(* IEC 61131-3 sources: daoli-st-library/DL_MathData (part 28) *)

(* ---- FC_DL_WordToBytes.st ---- *)
(*==============================================================================
 * 组件名称 (Component)  : FC_DL_WordToBytes
 * 所属子库 (Sublibrary) : DL_MathData
 * 当前版本 (Version)    : 1.0.0
 * 兼容性   (Platform)   : CODESYS 3.5 / TwinCAT 3 / 汇川 InoProShop / Machine Expert
 *                         仅依赖 Standard.library（SHR / AND / 类型转换），零厂商方言
 * 来源标签 (Source)     : t2-1-lgf-converter（字节序拆解族，clean-room 编写）
 * 功能描述 (Function)   : WORD / DWORD 按字节序拆解为 BYTE 数组（写经指针输出）。
 *                         槽位语义与 FC_DL_WordFromBytes 完全对偶：槽 0 = 最高字节；
 *                         映射为对合映射（ involutive），同一序号下
 *                         WordToBytes(WordFromBytes(bytes, eOrder, len), eOrder, len)
 *                         逐字节还原源数组（round-trip 验收）。
 *                         nValueLen = 2 时只取低 16 位（高 16 位忽略）。
 *                         缓冲长度不足时钳位只写前 nBufLen 个槽位并置信息级。
 * 归属声明 (Ownership)  : E_DL_ByteOrder 归属 DL_MathData\FC_DL_SwapBytes32.st，
 *                         本件只引用不重声明（FB51-7）。
 * 边界与语义披露 (Boundary disclosure) :
 *   1) 指针 NIL 或缓冲长度 <= 0：结构性早退，不写任何字节，返回 FALSE（零写入语义）。
 *   2) 缓冲长度大于目标长度：多余槽位不触碰（不置码——缓冲边界由调用方持有，
 *      可观测性在调用方，R90 反证成立不加码）。
 *   3) 还原方向不饱和（R81 披露）：本件是拆解不是还原时刻 / 标识，拆解失败
 *      返回 FALSE + 故障级码，绝无静默饱和写入。
 *   4) 移位量上界 (nLenUse-1-j)*8 结构性 <= 24 < 32（DWORD 位宽），禁 MOD 归一的
 *      不变量由本披露承担（R48 口径）。
 *   5) 验收向量（与 FromBytes 对拍）：CDAB 序 16#0000_1234 -> {16#34, 16#12}；
 *      ABCD 16#1234_5678 -> {16#12,16#34,16#56,16#78}；缓冲 1 字节拆 DWORD
 *      -> 只写最高字节 + 信息级钳位。
 * 故障码表 (Error codes) :
 *   16#0001_03F5 [故障级] 缓冲指针 NIL 或 nBufLen <= 0，不写任何字节，返回 FALSE
 *                 反证：未写缓冲与「缓冲区内容本来如此」不可区分（本件无权回读
 *                 调用方缓冲），码位是唯一的失败事实出口。
 *   16#0001_03F6 [故障级] 字节序枚举越界（非 0..3），回退默认大端 eAbcd 继续服务
 *                 反证：回退结果与显式填 eAbcd 输出组合相同，码位承载组态有误事实。
 *   16#0001_04BA [信息级] 缓冲长度不足目标长度，已钳位只写前段
 *                 反证：钳位写入与「调用方只想要前段」输出组合相同，无码不可区分。
 *   16#0001_04BB [信息级] nValueLen 非 2/4，回退默认 WORD（2 字节）继续服务
 *                 反证：回退结果与显式填 2 相同，码位承载组态有误事实。
 * 码位总账 (Code ledger) : 16#0001_03F5 / 03F6 用 ｜ 16#0001_04BA / 04BB 用
 * 依赖     (Depends)    : TYPE E_DL_ByteOrder（属主 FC_DL_SwapBytes32.st，只引用）
 * 红线自检 (Redline)    : R1 ✓ 零全局变量与 VAR_EXTERNAL ｜ R2 ✓ 零 %I/%Q 物理地址
 *                         R3 ✓ 纯 IEC 61131-3（指针判空 + 标准移位/转换）
 *                         R4 ✓ 指针 NIL 闸 / 缓冲域闸 / 枚举域闸 / 全分支码位配对
 *                         R5 ✓ 全变量中英双语同行注释 ｜ R6 N/A（纯函数，无状态机）
 *                         R7 N/A（无定时器 / 边沿实例）
 * 修订历史 (Revision)   :
 *   2026-11-22  v1.0.0  首版入库（R68 构建轮 · 批 1 · 目标 5）
 *============================================================================*)
FUNCTION FC_DL_WordToBytes : BOOL
VAR_INPUT
    uValue    : DWORD;              // 待拆解值（WORD 目标时只取低 16 位）/ Value to split, low word only for WORD
    nValueLen : INT := 2;           // 值长度 [字节]，2 = WORD，4 = DWORD / Value length in bytes
    eOrder    : E_DL_ByteOrder;     // 字节序选择（属主 FC_DL_SwapBytes32.st）/ Byte order selector
    nBufLen   : INT;                // 输出缓冲长度 [字节]，<= 0 无效 / Output buffer length, <= 0 invalid
    pBuf      : POINTER TO BYTE;    // 输出缓冲首指针（指针本身不被改写，按输入口径）/ Output buffer pointer, never re-pointed
END_VAR
VAR_OUTPUT
    bWritten  : BOOL;    // 本拍写入成功 / Write succeeded this call
    bError    : BOOL;    // 故障标志（0307 / 0308 置位，R45 配对）/ Fault flag, set on 0307 and 0308
    uInfoId   : UDINT;   // 故障码，0 = 无故障（纯函数每拍重算）/ Error code, recomputed per call
END_VAR
VAR
    nWriteLen : INT;     // 本拍实际写入字节数 [个] / Bytes actually written this call
    nSlotByte : INT;     // 当前槽位映射回的源字节下标 / Byte index the current slot maps back to
    nShift    : DINT;    // 当前槽位移位量 [bit]，结构性 <= 24 / Slot shift amount
    uSlotVal  : DWORD;   // 当前槽位值（已掩码低 8 位）/ Current slot value, low 8 bits
    uB        : BYTE;    // 当前槽位字节 / Current slot byte
    nLenUse   : INT;     // 钳位后的值长度 [字节] / Clamped value length
    bOrderOk  : BOOL;    // 字节序枚举合法性 / Byte order validity
    j         : INT;     // 槽位遍历索引 / Slot loop index
END_VAR
VAR CONSTANT
    DL_WTB_LEN_MIN : INT      := 2;          // 值长度下限 [字节]（WORD）/ Value length floor, WORD
    DL_WTB_LEN_MAX : INT      := 4;          // 值长度上限 [字节]（DWORD）/ Value length ceiling, DWORD
    DL_WTB_MASK_FF : DWORD    := 16#0000_00FF; // 低 8 位掩码 / Low byte mask
END_VAR

(*------------------------------------------------------------------------------
 * 段 1｜安全预置（P-01 范式）：任何异常路径不写缓冲、返回 FALSE
 *      Safe preset: every exceptional path writes nothing and returns FALSE
 *-----------------------------------------------------------------------------*)
FC_DL_WordToBytes := FALSE;
bWritten := FALSE;
bError   := FALSE;
uInfoId  := 16#0000_0000;

(*------------------------------------------------------------------------------
 * 段 2｜域闸（R151 全枚举：指针 + 缓冲 + 值长度 + 枚举四闸）
 *      Domain gates: pointer, buffer, value length and enum
 *-----------------------------------------------------------------------------*)
IF (pBuf = 0) OR (nBufLen <= 0) THEN
    uInfoId := 16#0001_03F5;    // 故障级：指针 NIL 或缓冲非法 / Fault: NIL pointer or bad buffer
    bError  := TRUE;            // R45 配对 / Paired with the fault code
    RETURN;                     // 结构性早退：输出已全预置，零写入语义成立（规格明示豁免）
END_IF

IF (nValueLen < DL_WTB_LEN_MIN) OR (nValueLen > DL_WTB_LEN_MAX) THEN
    nLenUse := DL_WTB_LEN_MIN;  // 二级回退：钳回默认 WORD（R117 两级参数回退）
    uInfoId := 16#0001_04BB;    // 信息级：值长度非法回默认 / Info: length defaulted
ELSE
    nLenUse := nValueLen;       // 合法直通 / Valid pass-through
END_IF

bOrderOk := (eOrder = E_DL_ByteOrder.eAbcd) OR (eOrder = E_DL_ByteOrder.eDcba)
            OR (eOrder = E_DL_ByteOrder.eBadc) OR (eOrder = E_DL_ByteOrder.eCdab);
IF NOT bOrderOk THEN
    uInfoId := 16#0001_03F6;    // 故障级：字节序越界回默认大端（0142 风格先例口径）/ Fault: order defaulted
    bError  := TRUE;            // R45 配对 / Paired with the fault code
END_IF

(*------------------------------------------------------------------------------
 * 段 3｜写入长度钳位（边界 B4）：缓冲不足只写前段 + 信息级
 *      Write length clamp: short buffer writes the leading slots only
 *-----------------------------------------------------------------------------*)
IF nBufLen < nLenUse THEN
    nWriteLen := nBufLen;       // 钳位：只写缓冲能容纳的槽位 / Clamp to buffer capacity
    uInfoId   := 16#0001_04BA;  // 信息级：缓冲不足钳位 / Info: buffer clamped
ELSE
    nWriteLen := nLenUse;       // 充足：全量写入 / Full write
END_IF

(*------------------------------------------------------------------------------
 * 段 4｜拆解主体（边界 B1/B3）：取槽 -> 掩码 -> 降位 -> 反映射 -> 写缓冲
 *      Split body: slot, mask, narrow, inverse-map, write buffer
 *      反映射即对合映射本身：i = map(j)（映射自逆，与 FromBytes 同口径）
 *-----------------------------------------------------------------------------*)
FOR j := 0 TO (nWriteLen - 1) DO
    (* 槽位到源字节下标的对合映射（与 FromBytes 逐分支一致） *)
    (* Involutive slot to byte mapping, branch-aligned with WordFromBytes *)
    IF eOrder = E_DL_ByteOrder.eDcba THEN
        nSlotByte := (nLenUse - 1) - j;          // 全反序 / Full reverse
    ELSIF eOrder = E_DL_ByteOrder.eBadc THEN
        nSlotByte := (j XOR 1) MOD nLenUse;      // 寄存器内两两互换 / Swap within register pairs
    ELSIF eOrder = E_DL_ByteOrder.eCdab THEN
        IF nLenUse = DL_WTB_LEN_MAX THEN
            nSlotByte := (j XOR 2) MOD nLenUse;  // DWORD：高低字互换 / DWORD: word swap
        ELSE
            nSlotByte := 1 - j;                  // WORD：退化为字节反序（见头披露）/ WORD: degenerate reverse
        END_IF
    ELSE
        nSlotByte := j;                          // eAbcd 大端直排（含越界回退默认）/ Big endian, incl. fallback
    END_IF

    nShift   := (nLenUse - 1 - j) * 8;                   // 槽位移位量，结构性 <= 24 / Slot shift
    uSlotVal := SHR(uValue, nShift) AND DL_WTB_MASK_FF;  // 取槽位并掩低 8 位 / Slot value masked
    uB       := DWORD_TO_BYTE(uSlotVal);                 // 降位到字节 / Narrow to byte
    pBuf[nSlotByte] := uB;                               // 反映射写入缓冲 / Inverse-mapped write
END_FOR

(*------------------------------------------------------------------------------
 * 段 5｜结果回写：全量或钳位写入均算成功（钳位事实由 0409 承载）
 *      Result write-back: full or clamped write both count as success
 *-----------------------------------------------------------------------------*)
FC_DL_WordToBytes := TRUE;
bWritten := TRUE;
END_FUNCTION

(* ---- FC_DL_WordToIntSat.st ---- *)
(*
    FC_DL_WordToIntSat —— WORD 到 INT 的双语义落地
    ------------------------------------------------------------------
    分类      : DL_MathData / Convert
    前缀      : FC_DL_
    版本      : 1.0.0
    溯源      : IEC 61131-3 标准语义的道莅防御性实现（WORD 16 位无符号 → INT 16 位有符号）；
                域内委托平台内建 WORD_TO_INT，本件不重实现数学内核；
                补码解释偏移量、饱和出口、双语义开关、错误分级与码位 100% 自有；
                clean-room 重写，未复制任何闭源厂商源码，参考实现仅限 MIT/Apache 许可
    平台      : 纯 IEC 61131-3，CODESYS V3.5+ / TwinCAT 3 / InoProShop 通用
    作者      : 道莅代码库 · PLC编程专家（R20）
    ------------------------------------------------------------------
    功能说明  : Modbus 16 位寄存器搬上来的是无符号位型，落到 INT 工程量时现场存在两种合法口径：
                ① 补码解释——仪表把 −200~−1 的工程量以 65336~65535 的补码形式放在寄存器里，
                   直接截成 INT 就得到 −200 是正确的，此时「饱和到 32767」反而是错的；
                ② 上饱和——纯正计数/量程值，超 32767 只能钳位。
                两种口径业务含义完全相反，靠猜必错，故本件用显式引脚 bTwosComplement 由调用方声明，
                并把「发生了哪一种」用 bInterpreted 回告，HMI 与追责链都看得见。
                核心防御：① 补码解释全程在 DINT 域做减法（升位后再减 65536），
                   禁在 INT 域内做减法——16 位域内减法中途溢出是三平台回绕差异的经典源头；
                ② 域内直接委托内建，零额外开销；
                ③ 三种出路（原值 / 补码 / 饱和）都是安全侧取值，值本身仍可用，
                   故本件故障级三槽全预留，只在信息级区分口径。
                职责边界：DWORD 降位归 FC_DL_DwordToIntSat，LWORD 降位归
                FC_DL_LwordToLintSat；本件只管 16 位双语义。
    编译门槛  : 主路径依赖平台内建 WORD_TO_INT / WORD_TO_DINT / DINT_TO_INT，
                均为 IEC 61131-3 标准转换函数，三平台标准库均提供，无厂商方言。
    错误码    : 16#0001_0416 超域且按补码解释为负值（已升 DINT 再减偏置）——信息级，值可用
                16#0001_0417 超域且按上饱和处理（钳位至 32767）——信息级，值可用
                16#0001_033F 预留（故障级，不得挪用）
                16#0001_0340 预留（故障级，不得挪用）
                16#0001_0341 预留（故障级，不得挪用）
    码位总账  : 16#0001_0416 用 / 16#0001_0417 用 ｜ 16#0001_033F 预留 / 16#0001_0340 预留 / 16#0001_0341 预留
    状态机    : R6 标注 N/A —— 本组件为纯函数无顺序状态机，无 CASE 可写，非法状态不可能出现
    采样约定  : 本件无定时器、无沿检测、无状态；单拍纯计算，结论与任务周期无关。
    修订记录  : 2026-11-16 v1.0.0 首次入库（R20）
*)
FUNCTION FC_DL_WordToIntSat : INT
VAR_INPUT
    uIn              : WORD;                  // 输入值 [无量纲]，全域 0~65535 / input value [dimensionless], full WORD domain
    bTwosComplement  : BOOL := FALSE;         // TRUE = 超域按补码解释为负值；FALSE = 上饱和至 32767 / TRUE interprets the overrun as two's complement, FALSE saturates
END_VAR
VAR_OUTPUT
    eErr             : UDINT;                 // 错误码，0=正常 / error id, 0=ok
    bError           : BOOL;                  // 故障标志，本件无故障级出口，恒为 FALSE / error flag, always FALSE here as no fault exit exists
    bValid           : BOOL;                  // 返回值是否可用（三种出路均可用）/ return usable, all three exits are usable
    bInterpreted     : BOOL;                  // 发生了补码解释或上饱和 / a two's complement interpretation or a saturation happened
END_VAR
VAR CONSTANT
    DL_INT_MAX_AS_WORD : WORD := 32767;       // INT 上限的 WORD 形态 [无量纲] / the INT maximum expressed as WORD [dimensionless]
    DL_INT_MAX       : INT := 32767;          // INT 上限值 [无量纲] / the INT maximum value [dimensionless]
    DL_INT_ZERO      : INT := 0;              // 有符号零常量，避免裸字面量 [无量纲] / signed zero constant [dimensionless]
    DL_TWOS_BIAS     : DINT := 65536;         // 补码解释偏移量，即 2^16 [无量纲] / two's complement bias, 2 to the 16 [dimensionless]
END_VAR
VAR
    nTmp             : DINT;                  // 补码解释中间量，先升 DINT 再减 [无量纲] / two's complement intermediate, widened before subtracting [dimensionless]
    nOut             : INT;                   // 结果中间量 [无量纲] / result intermediate [dimensionless]
END_VAR

// 段 1｜返回值与错误状态预置 / segment 1, preset return value and error status
FC_DL_WordToIntSat := DL_INT_ZERO;            // 故障缺省返回 0 [无量纲] / fault default returns zero [dimensionless]
eErr := 0;                                    // 预置无错误 / preset no error
bError := FALSE;                              // 本件无故障级出口，恒 FALSE / no fault exit exists, always FALSE
bValid := FALSE;                              // 预置不可用，通过闸门后置位 / preset invalid, set TRUE after the gates
bInterpreted := FALSE;                        // 预置未做解释或饱和 / preset no interpretation and no saturation
nOut := DL_INT_ZERO;                          // 结果中间量清零 / clear the result intermediate

// 段 2｜域内闸：不超过 32767 即零开销直通 / segment 2, in-domain gate, zero overhead pass-through
IF uIn <= DL_INT_MAX_AS_WORD THEN
    nOut := WORD_TO_INT(uIn);                 // 域内委托内建 [无量纲] / in-domain delegation to the built-in [dimensionless]
    bValid := TRUE;                           // 直通值可用 / the pass-through value is usable
ELSE
    // 段 3｜超域双语义分派（口径由调用方显式声明，绝不猜测）/ segment 3, explicit dual-semantics dispatch
    IF bTwosComplement THEN
        nTmp := WORD_TO_DINT(uIn) - DL_TWOS_BIAS; // 先升 DINT 再减偏置，禁在 INT 域内减法 / widen to DINT before subtracting, never subtract inside INT
        nOut := DINT_TO_INT(nTmp);            // 结果已在 −32768~−1，回转 INT 无损 / the result is already inside −32768 to −1, the narrowing is lossless
        bInterpreted := TRUE;                 // 标记已做补码解释 / flag the two's complement interpretation
        eErr := 16#0001_0416;                 // 信息级：超域按补码解释为负值 / info level, the overrun was read as two's complement
    ELSE
        nOut := DL_INT_MAX;                   // 上饱和至 32767 / saturate to the INT maximum
        bInterpreted := TRUE;                 // 标记已做上饱和 / flag the saturation
        eErr := 16#0001_0417;                 // 信息级：超域已饱和，值仍可用 / info level, saturated, still usable
    END_IF
    bValid := TRUE;                           // 两种出路都是安全侧取值 / both exits stay on the safe side
END_IF

// 段 4｜发布结果 / segment 4, publish the result
FC_DL_WordToIntSat := nOut;                   // 输出 16 位有符号结果 [无量纲] / publish the signed 16-bit result [dimensionless]
bError := FALSE;                              // 信息级不置故障（双保险）/ info level never raises a fault, second line of defence
END_FUNCTION

(* ---- FC_DL_WrapAngleDeg.st ---- *)
(*
    组件名称 : FC_DL_WrapAngleDeg
    所属子库 : DL_MathData
    当前版本 : 1.0.0
    兼 容 性 : CODESYS V3.5+ / TwinCAT 3 / 汇川 InoProShop；仅依赖 Standard.library
    功能描述 : 角度归一原子，把任意角度折算到 (−180, 180]（缺省）或 [0, 360)，并顺带出口圈数供多圈相位追溯。
              取舍 ①：禁 MOD —— REAL/LREAL 上的 MOD 在三平台上的「余数符号」与「负零」行为不一致，
              而且 MOD 结果可能给出 -0.0 与 360.0 两种等价表示，会让下游的相等判据抖动。
              本件改用「TRUNC 求整圈数 + 一次条件加减」，最多一次加减即可落到目标半开区间。
              取舍 ②：超可归一域直接报故障而不钳位 —— 角度钳位会静默改变转向语义（-720° 被钳成 -180°
              就成了反向），运动链上这是灾难；宁可停机让调用方查清输入来源。
              取舍 ③：零容差归一为 +0.0 —— 消除 -0.0 与「恰好 360.0」两种抖动值，让下游可以用符号判方向。
              取舍 ④：DL_GUARD_MAX 仅作防御性预留常量而非死代码 —— 本实现全文无循环（条件加减最多一次），
              守卫计数器无使用场景；保留该常量是为了在扩展为多圈归一时有现成的上限口径，
              避免届时再引入裸数值。此处显式留档，不留未解释常量。
    开源溯源 : 原创实现。运动层 CamPhaseTrim / ElectronicCam 反复手写同一段归一并多次留痕，；本件为 IEC 61131-3 标准语义的道莅防御性实现（原创实现，零外部源码复制）。
              本件为其唯一原子出口。无外部源码参考，码位与分级 100% 自有。
    本文件内含 : FUNCTION FC_DL_WrapAngleDeg（单 POU，无配套类型）
    依 赖 : 无 DL_ 内部依赖；Standard.library: 无
    红线自检 : R1 ✓ 零全局变量与外部变量 ｜ R2 ✓ 零物理 IO 地址
              R3 ✓ 纯 IEC 61131-3 ｜ R4 ✓ 非有限闸 + 可归一域闸 + 零容差归一（禁 MOD、禁循环、禁钳位）
              R5 ✓ 全变量中英双语同行注释 ｜ R6 N/A 纯函数无顺序状态机，无 CASE 可写
              R7 N/A 无定时器、无沿检测实例 ｜ R8 ✓ 全部域与容差常量化（含守卫常量用途说明）
    错误码   : 16#0001_043C [信息级] 输入超一圈已归一，bValid = TRUE
               16#0001_043D [信息级] 结果落零容差已归一为 +0.0，bValid = TRUE
               16#0001_0378 [故障级] 输入非有限（NaN 或 ±INF），返回 0，bValid = FALSE
               16#0001_0379 [故障级] 超可归一域（|角度| > DL_ANGLE_ABS_MAX），返回 0，bValid = FALSE
               16#0001_037A [故障级] 预留禁用（不得挪用）
    码位总账 : 16#0001_043C 用 / 16#0001_043D 用 ｜ 16#0001_0378 用 / 16#0001_0379 用 / 16#0001_037A 预留
    遗留假设 : ① LREAL_TO_DINT 对超出 DINT 域的输入行为未定义，本件已用 DL_ANGLE_ABS_MAX = 1E6 把商限制在 ±2778，
              结构性不进该分支；该上限本身为推导，未三平台实测。
              ② TRUNC 返回值宽度与入参一致（LREAL），用于 LREAL_TO_DINT 前置 —— IEC 语义推导，未逐平台实测。
    修订历史 :
        2026-11-16  v1.0.0  首版，R21 批次 1 入库
*)
FUNCTION FC_DL_WrapAngleDeg : LREAL
VAR_INPUT
    fAngleDeg       : LREAL := 0.0;   // 任意角度，有效域 |x| ≤ 1E6 [°] / arbitrary angle, valid up to one million degrees [deg]
    bZeroTo360      : BOOL := FALSE;  // FALSE → (−180, 180]；TRUE → [0, 360) / FALSE gives minus 180 to 180, TRUE gives zero to 360 [range]
END_VAR
VAR_OUTPUT
    eErr            : UDINT;          // 错误码，0=正常；16#0001_04XX 信息级 / 16#0001_03XX 故障级 / error id, 0=ok
    bError          : BOOL;           // 故障级标志，eErr 落 16#0001_03XX 时为 TRUE / fault flag, TRUE on fault-level eErr
    bValid          : BOOL;           // 归一结果是否可用 / normalised result usable flag
    nTurns          : DINT;           // 圈数，向零取整，供多圈相位追溯 [圈] / completed turns truncated toward zero, for multi-turn phase tracing [turn]
END_VAR
VAR
    fQuot           : LREAL;          // 角 / 360 的商 [圈] / quotient of the angle over one turn [turn]
    fRet            : LREAL;          // 归一结果工作寄存器 [°] / normalisation working register [deg]
    bOverOneTurn    : BOOL;           // 输入绝对值是否已超一圈 / whether the magnitude already exceeds one turn
END_VAR
VAR CONSTANT
    DL_DEG_PER_TURN     : LREAL := 360.0;                      // 一圈的角度 [°] / degrees per turn [deg]
    DL_DEG_HALF_TURN    : LREAL := 180.0;                      // 半圈，区间判定边界 [°] / half turn, the interval boundary [deg]
    DL_ANGLE_ABS_MAX    : LREAL := 1.0E6;                      // 可归一域上限，超此值 LREAL 已无 0.001° 分辨率 [°] / normalisable domain limit [deg]
    DL_FLOAT_EPS        : LREAL := 1.0E-9;                     // 零容差，比 0.001° 分辨率小两个量级 [°] / zero tolerance, two decades below the resolution [deg]
    DL_LREAL_MAX_FINITE : LREAL := 1.7976931348623157E308;     // LREAL 最大有限值 [无量纲] / largest finite LREAL [dimensionless]
    DL_LREAL_ZERO       : LREAL := 0.0;                        // 零哨兵，归一目标值 [无量纲] / zero sentinel and normalisation target [dimensionless]
    DL_GUARD_MAX        : DINT := 1000;                        // 守卫上限预留（本件无循环，见头注释取舍 ④）[次] / reserved guard limit, unused here because there is no loop [count]
    DL_ERR_NONE         : UDINT := 16#0000_0000;               // 无故障 / no error
END_VAR

// 段 1｜返回值与错误状态预置 / segment 1, preset the return value and the error state
FC_DL_WrapAngleDeg := DL_LREAL_ZERO;    // 故障缺省返回 0 / fault default returns zero
eErr   := DL_ERR_NONE;                  // 预置无错误 / preset no error
bError := FALSE;                        // 预置无故障 / preset no fault
bValid := FALSE;                        // 预置结果不可用 / preset unusable
nTurns := 0;                            // 预置圈数 0 / preset the turn count to zero

// 段 2｜输入有限性闸 / segment 2, input finiteness gate
IF (fAngleDeg <> fAngleDeg) OR (ABS(fAngleDeg) > DL_LREAL_MAX_FINITE) THEN
    eErr   := 16#0001_0378;             // 输入非有限（故障级）/ non-finite input, fault level
    bError := TRUE;                     // 置故障标志 / raise the fault flag
    RETURN;                             // 返回 0，bValid 保持 FALSE / return zero, bValid stays FALSE
END_IF

// 段 3｜可归一域闸：超域不钳位，钳位会静默改转向 / segment 3, domain gate, clamping would silently flip the direction
IF ABS(fAngleDeg) > DL_ANGLE_ABS_MAX THEN
    eErr   := 16#0001_0379;             // 超可归一域（故障级）/ beyond the normalisable domain, fault level
    bError := TRUE;                     // 置故障标志 / raise the fault flag
    RETURN;                             // 返回 0，bValid 保持 FALSE / return zero, bValid stays FALSE
END_IF

// 段 4｜整圈剥离：TRUNC 求圈数，再一次性减掉，禁 MOD / segment 4, whole turns stripped with TRUNC, never with MOD
fQuot  := fAngleDeg / DL_DEG_PER_TURN;                                  // 商，域内 |商| ≤ 2778，转换结构性安全 / the quotient stays within plus or minus 2778 by construction
nTurns := LREAL_TO_DINT(TRUNC(fQuot));                                  // 向零取整得圈数 / truncate toward zero to get the turns
fRet   := fAngleDeg - DINT_TO_LREAL(nTurns) * DL_DEG_PER_TURN;          // 剥离整圈后的余量，落在 (−360, 360) / the remainder after stripping whole turns
bOverOneTurn := ABS(fAngleDeg) > DL_DEG_PER_TURN;                       // 记录「曾超一圈」/ remember that the input exceeded one turn

// 段 5｜一次条件加减落到目标半开区间（最多一次，不写循环）/ segment 5, one conditional add or subtract at most
IF fRet > DL_DEG_HALF_TURN THEN
    fRet := fRet - DL_DEG_PER_TURN;     // 上半圈搬下来 / bring the upper half down
ELSIF fRet <= -DL_DEG_HALF_TURN THEN
    fRet := fRet + DL_DEG_PER_TURN;     // 下半圈搬上去，(-180] 边界归 +180 / bring the lower half up, the boundary joins plus 180
END_IF

// 段 6｜零容差归一：消除 −0.0 与 360.0 抖动 / segment 6, zero tolerance normalisation removes minus zero and 360 jitter
IF ABS(fRet) < DL_FLOAT_EPS THEN
    fRet := DL_LREAL_ZERO;              // 一律归 +0.0 / always normalise to positive zero
    eErr := 16#0001_043D;               // 零容差归一（信息级，不置 bError）/ zero tolerance hit, info level
END_IF

// 段 7｜区间搬移：0..360 口径 / segment 7, shift into the zero to 360 interval when requested
IF bZeroTo360 THEN
    IF fRet < DL_LREAL_ZERO THEN
        fRet := fRet + DL_DEG_PER_TURN; // 负半区搬到正半区，结果恒 < 360 / move the negative half up, the result stays below 360
    END_IF
END_IF

// 段 8｜超一圈提示（先置者保留原则：043C 若已被占则不覆盖）/ segment 8, one-turn hint, never overwriting an existing code
IF bOverOneTurn AND (eErr = DL_ERR_NONE) THEN
    eErr := 16#0001_043C;               // 输入超一圈已归一（信息级）/ input beyond one turn, info level
END_IF

// 段 9｜出口 / segment 9, exit
FC_DL_WrapAngleDeg := fRet;             // 输出归一角度 / publish the normalised angle
bValid := TRUE;                         // 结果可用 / the result is usable
END_FUNCTION

(* ---- FC_DL_WrapAngleNorm.st ---- *)
// FC_DL_WrapAngleNorm v1.0.0
(*==============================================================================
 * 功能描述: 角度归一化到 [-180, 180) 区间。fmod 风格两段修正：先以 TRUNC 取整
 *           折返 (-360,360)，再单侧修正进 [-180,180)；非有限输入返回 0 并置
 *           bValid=FALSE。同名避让：库内已有 FC_DL_WrapAngleDeg。
 * 接口契约: 输入 fAngleDeg [°]；输出 bValid 回执，返回归一后角度 [°]。
 * 修订历史: 2026-11-23  v1.0.0  R74 首版
 *==============================================================================*)

FUNCTION FC_DL_WrapAngleNorm : REAL
VAR_INPUT
    fAngleDeg : REAL := 0.0;   // 输入角度（任意域）[°] / Input angle, any range [deg]
END_VAR
VAR_OUTPUT
    bValid : BOOL;             // 结果有效回执 [-] / Result validity receipt
END_VAR
VAR
    fW : REAL;                 // 折返工作角 [°] / Folded working angle
END_VAR

(* —— 段 0：全路径赋值缺省（无效安全侧） —— *)
bValid := FALSE;                             // 有效回执预清 / Validity preset
FC_DL_WrapAngleNorm := 0.0;                  // 返回角缺省零 / Result default zero

(* —— 段 1：非有限与幅值闸（NaN 自反判 + 近 Inf 兜底） —— *)
IF fAngleDeg <> fAngleDeg THEN               // NaN 自反判（判等禁令唯一例外） / NaN self-reflexive test
    RETURN;                                  // 无效返回零 / Invalid, return zero
END_IF
IF ABS(fAngleDeg) >= 1.0E15 THEN             // 近 Inf 幅值闸（TRUNC 精度域兜底） / Near-Inf magnitude gate
    RETURN;                                  // 无效返回零 / Invalid, return zero
END_IF

(* —— 段 2：两段归一化（TRUNC 折返 → 单侧修正进 [-180,180)） —— *)
fW := fAngleDeg - 360.0 * TRUNC(fAngleDeg / 360.0);   // 第一段：折返到 (-360,360) / First fold into (-360,360)
IF fW >= 180.0 THEN                          // 第二段：上界修正进 [-180,180) / Upper correction into range
    fW := fW - 360.0;
ELSIF fW < -180.0 THEN                       // 第二段：下界修正进 [-180,180) / Lower correction into range
    fW := fW + 360.0;
END_IF
FC_DL_WrapAngleNorm := fW;                   // 返回归一后角度 / Return wrapped angle
bValid := TRUE;                              // 有效回执 / Validity receipt

END_FUNCTION

(* ---- FC_DL_WrapIndexNeg.st ---- *)
(*
  Name        : FC_DL_WrapIndexNeg
  Category    : DL_MathData
  Version     : 1.0.0
  Purpose     : 环窗下标负值模归正：把任意（含负）下标折叠进 [1..N] 或 [0..N-1] 合法区间，修正 IEC MOD 负余数语义；/ Fold any index (negative allowed) into [1..N] or [0..N-1], correcting IEC MOD negative-remainder semantics
  溯源        : 自研·环窗族治理（R193 配套），IEC 61131-3 标准语义的道莅防御性实现
  Boundary    : ① 模基数 diMod <= 0 → 返回 0 哨兵，不做除法（防除零）；
                ② IEC MOD 余数符号随被除数（负被除数得负余数），本件统一 +diMod 归正一次；
                ③ 1 基口径下 (diIdx - 1) 有下溢风险，先钳到 DINT 可表区间再折算；
                ④ 纯整型运算，无浮点比较、无 NaN/Inf 路径。
*)
FUNCTION FC_DL_WrapIndexNeg : DINT
VAR_INPUT
    diIdx     : DINT := 0;                   (* 输入下标，允许负值（如倒序回看 -3 表示前 3 个）[-] / Input index, negative allowed *)
    diMod     : DINT := 1;                   (* 模基数（窗深/表长），域 > 0 [-] / Modulus base, must be > 0 *)
    xOneBased : BOOL := TRUE;                 (* TRUE = 1 基口径 [1..diMod]；FALSE = 0 基口径 [0..diMod-1] [-] / 1-based or 0-based *)
END_VAR
VAR
    diBase : DINT;                            (* 折算到 0 基的中间量 [-] / Value folded to 0-based *)
    diRem  : DINT;                            (* IEC MOD 余数（可负，须归正）[-] / IEC MOD remainder, may be negative *)
END_VAR
VAR CONSTANT
    DL_WIN_DINTMAX : DINT := 2147483647;      (* DINT 可表上限（折算前钳位基准，R28 双边界）[#] / DINT representable max *)
    DL_WIN_DINTMIN : DINT := -2147483647;     (* 安全下限（避开 -2^31 取负溢出的自反陷阱）[#] / Safe DINT min avoiding negation overflow *)
END_VAR

(* —— 段 1：模基数闸（除零与非法基数唯一出入口，返回哨兵 0） —— *)
IF diMod <= 0 THEN
    FC_DL_WrapIndexNeg := 0;                  (* 哨兵 0：调用侧须以 diMod 闸先行拒绝 / Sentinel 0, caller must gate diMod *)
    RETURN;
END_IF

(* —— 段 2：输入下标双侧钳位（防 -2^31 取负溢出与 1 基折算下溢） —— *)
IF diIdx > DL_WIN_DINTMAX THEN
    diIdx := DL_WIN_DINTMAX;                  (* 上限钳位（可表性反算，非饱和业务语义） / Upper clamp for representability *)
ELSIF diIdx < DL_WIN_DINTMIN THEN
    diIdx := DL_WIN_DINTMIN;                  (* 下限钳位（-2^31 不参与折算，避开自反溢出） / Lower clamp avoiding self-negation overflow *)
END_IF

(* —— 段 3：折算到 0 基 + 负余数归正 —— *)
IF xOneBased THEN
    diBase := diIdx - 1;                      (* 1 基 → 0 基（已钳位，无下溢） / 1-based to 0-based *)
ELSE
    diBase := diIdx;                          (* 0 基直接用 / 0-based direct *)
END_IF
diRem := diBase MOD diMod;                    (* IEC MOD：余数符号随被除数，负被除数得负余数 / IEC MOD keeps dividend sign *)
IF diRem < 0 THEN
    diRem := diRem + diMod;                   (* 归正一次即落入 [0, diMod-1]（|diRem| < diMod 保证一次足够） / One fold suffices *)
END_IF

(* —— 段 4：回写目标口径 —— *)
IF xOneBased THEN
    FC_DL_WrapIndexNeg := diRem + 1;          (* 0 基 → 1 基，域 [1..diMod] / Back to 1-based *)
ELSE
    FC_DL_WrapIndexNeg := diRem;              (* 0 基直接输出，域 [0..diMod-1] / 0-based output *)
END_IF
END_FUNCTION

(* ---- FC_DL_YarnCountConvert.st ---- *)
(*
  DL Factory R83 | FC_DL_YarnCountConvert
  功能：在棉英制支数 Ne、公制支数 Nm、特数 Tex、旦尼尔 Den 之间双向换算。
  开源溯源：无（clean-room 自研，依据公开工艺公式，来源=行业通用公式，许可证=MIT，借鉴点=公式结构）
  规则：R1-R21 全遵守
*)
FUNCTION FC_DL_YarnCountConvert : REAL
VAR_INPUT
    fCount   : REAL; // 输入支数值（须为正）[-] / Input count value, positive [-]
    iFromSys : INT;  // 源制式 1=Ne 2=Nm 3=Tex 4=Den / Source system code
    iToSys   : INT;  // 目标制式 1=Ne 2=Nm 3=Tex 4=Den / Target system code
    fDensity : REAL; // 纤维密度（量纲自检用）[g/cm³] / Fibre density for dimension check
END_VAR
VAR_OUTPUT
    fTexOut   : REAL; // 中间基准特数 [tex = g/1000m] / Intermediate linear density [tex]
    fCountOut : REAL; // 目标制式支数值 [-]/ Converted count in target system [-]
    xValid    : BOOL; // 计算有效性标志 / Calculation validity flag
END_VAR
VAR
    fTex : REAL; // 基准特数中间量 [tex] / Intermediate tex value [tex]
END_VAR
fTexOut := 0.0; fCountOut := 0.0; xValid := FALSE;  // 出口预置（R256）
// 非有限拦截 + 制式码域闸 + 密度量纲自检（R20/R21）
IF NOT (fCount > -1.0E30 AND fCount < 1.0E30) OR NOT (fDensity > -1.0E30 AND fDensity < 1.0E30) OR fCount <= 0.0 OR iFromSys < 1 OR iFromSys > 4 OR iToSys < 1 OR iToSys > 4 OR fDensity <= 0.0 OR fDensity > 3.0 THEN
    FC_DL_YarnCountConvert := -1.0; RETURN;   // 哨兵 -1：支数非正、制式码或密度越界 / Sentinel -1
END_IF
// 第一段：源制式 → 基准特数 Tex（全部除式分母为 fCount，上面已判正）
IF iFromSys = 1 THEN
    fTex := 590.5 / fCount;         // 棉英制 Ne → Tex [tex] / Ne to tex
ELSIF iFromSys = 2 THEN
    fTex := 1000.0 / fCount;        // 公制支数 Nm → Tex [tex] / Nm to tex
ELSIF iFromSys = 3 THEN
    fTex := fCount;                 // 特数直通 [tex] / Tex passes through
ELSE
    fTex := fCount / 9.0;           // 旦尼尔 Den → Tex [tex] / Den to tex
END_IF
// 第二段：基准特数 Tex → 目标制式（fTex 由第一段保证为正，除法安全）
IF iToSys = 1 THEN
    fCountOut := 590.5 / fTex;      // Tex → 棉英制 Ne [-]/ Tex to Ne
ELSIF iToSys = 2 THEN
    fCountOut := 1000.0 / fTex;     // Tex → 公制支数 Nm [-]/ Tex to Nm
ELSIF iToSys = 3 THEN
    fCountOut := fTex;              // 特数直通 [-]/ Tex passes through
ELSE
    fCountOut := fTex * 9.0;        // Tex → 旦尼尔 Den [-]/ Tex to Den
END_IF
// 出口：正特数才视为有效，非正走故障缺省
IF fTex > 0.0 THEN fTexOut := fTex; xValid := TRUE; END_IF  // 输出基准特数并置有效 [tex]
FC_DL_YarnCountConvert := fCountOut; // 返回目标制式支数 [-]/ Return converted count [-]
END_FUNCTION

(* ---- FB_DL_DataResampler.st ---- *)
(*
  ==================================================================
  组件名 Component  : FB_DL_DataResampler
  分类   Category   : DL_MathData
  复杂度 Complexity  : 中
  版本   Version    : 1.0.0
  功能   Purpose    : 变周期数据重采样。新周期沿（bNewCycle 上升沿）锁存新
                      样本进双缓冲（fPrev/fLast），拍间按相位 fFrac ∈ [0,1]
                      线性插值桥接输出；周期缺口超 tGapMax 计丢拍 nLostCnt；
                      非有限样本拒收计数 nSkipCnt 并置 bBad（禁静默吞）。
                      测量评估族语义，与 FB_DL_MovingAverage 窗口滤波分工。
  来源   Source     : T2-1-lgf-measurement（测量评估族待挖项）
  溯源   Origin     : 周期沿锁存 + 线性插值桥接为公开工程语义，clean-room
                      自研实现，未复制 LGF 或任何厂商私有库源码。
  平台   Platform   : 纯 IEC 61131-3（Standard.library: TON / R_TRIG，无私有库）
  分工声明 Split     : 与 FB_DL_MovingAverage 分工——后者做窗口均值滤波，
                      本件做变周期样本锁存与拍间插值桥接。
  作者   Author     : 道莅代码库 · PLC 编程专家（R59）
  ------------------------------------------------------------------
  边界 Boundary     :
                      一 安全语义：样本不足两帧或末帧非有限时 fOut 安全侧
                         零、bValid 假（插值桥不外推）；
                      二 fFrac 越域 [0,1] 回夹并置 bClamped（信息级，单点
                         回夹防多处覆盖）；
                      三 缺口窗 tGapMax 到期单拍计丢拍一次（自复位窗，R188），
                         窗口末退出迁移（本库纪律④）；
                      四 非有限样本：环不写入、bBad 置位、nSkipCnt 计数
                         （本库纪律②）；
                      五 定时器与沿检测全部段 0 无条件周期刷新（R7）；
                      六 无全局变量、无外部变量声明、无物理地址寻址。
  修订记录 Revision  :
    2026-11-21  v1.0.0  R59 首版（批 2 · 序号 8）
  ==================================================================
*)

FUNCTION_BLOCK FB_DL_DataResampler
VAR_INPUT
    fIn       : LREAL := 0.0;  // 样本输入 [工程单位] / the sample input [engineering unit]
    bNewCycle : BOOL := FALSE; // 新周期标志，上升沿锁存样本 [-] / the new cycle flag, the rising edge latches the sample
    fFrac     : LREAL := 0.0;  // 插值相位，域 [0,1] [无量纲] / the interpolation phase, zero through one
    tGapMax   : TIME := T#5S;  // 周期缺口看门狗窗 [毫秒] / the cycle gap watchdog [millisecond]
    bEnable   : BOOL := TRUE;  // 使能，失能输出安全侧零 [-] / the enable, disabling zeroes the output
END_VAR
VAR_OUTPUT
    fOut     : LREAL := 0.0;  // 插值桥接输出 [工程单位] / the interpolated bridge outlet [engineering unit]
    bValid   : BOOL := FALSE; // 输出可用标志（双帧齐且有限）[-] / the output usable flag
    bClamped : BOOL := FALSE; // 相位回夹发生（信息级）[-] / the phase clamp happened, informational
    bBad     : BOOL := FALSE; // 非有限样本拒收实时标志 [-] / the non finite sample rejection flag
    nLostCnt : UDINT := 0;    // 丢拍计数 [拍] / the lost cycle count
    nSkipCnt : UDINT := 0;   // 非有限拒收计数 [次] / the skipped non finite count
END_VAR
VAR CONSTANT
    DL_DRS_CNTMAX : UDINT := 4294967294; // 计数防回绕上界 [次] / the counter anti wrap clamp bound
END_VAR
VAR
    _bInit  : BOOL := FALSE; // 首拍初始化标志（R310，真实使用：首拍安全态预置）/ the first scan flag, real use
    _fPrev  : LREAL := 0.0;  // 前帧锁存副本 [工程单位] / the previous latched sample copy
    _fLast  : LREAL := 0.0;  // 末帧锁存副本 [工程单位] / the last latched sample copy
    _bHave  : BOOL := FALSE; // 双帧齐备锁存 [-] / the two samples ready latch
    _bFin   : BOOL;          // 样本有限工作量 [-] / the sample finiteness work flag
    rtNew   : R_TRIG;        // 新周期沿检测，段 0 无条件刷新 / the new cycle edge, refreshed unconditionally
    tonGap  : TON;           // 缺口看门狗（自复位窗），段 0 无条件刷新 / the gap watchdog, the self reset window
END_VAR

// 段 0｜定时器与沿检测无条件周期刷新（禁入分支，R7）/ segment 0, the unconditional refresh
rtNew(CLK := bNewCycle); // 新周期沿 / the new cycle edge
tonGap(IN := bEnable AND (NOT rtNew.Q) AND (NOT tonGap.Q), PT := tGapMax); // 自复位缺口窗（R188：IN 串 NOT Q）/ the self reset gap window

// 段 1｜首拍初始化（R310 真实使用路径）：输出安全态显式预置 / segment 1, the first scan init, the safe preset
IF NOT _bInit THEN // 首拍一拍 / the first scan
    _bInit := TRUE; // 置首拍标志 / raise the flag
    fOut := 0.0; // 输出强制安全零 / force the safe zero
    bValid := FALSE; // 有效强制假 / force the valid false
END_IF

// 段 2｜丢拍计数（缺口窗到期单拍一次，窗口末退出迁移，边界三）/ segment 2, the lost cycle count
IF tonGap.Q THEN // 缺口窗到期（本拍为超窗第一拍）/ the gap window expired, the first scan beyond
    IF nLostCnt < DL_DRS_CNTMAX THEN // 计数防回绕 / the wrap guard
        nLostCnt := nLostCnt + 1; // 计丢拍一次 / count one lost cycle
    END_IF
END_IF

// 段 3｜新周期沿锁存（有限样本才入双缓冲，边界四）/ segment 3, the edge latch
_bFin := (fIn = fIn) AND ((fIn - fIn) = (fIn - fIn)); // 样本有限双判据（R79）/ the finiteness dual verdicts
IF rtNew.Q THEN // 新周期沿 / the new cycle edge
    IF _bFin THEN // 有限样本受理 / a finite sample accepted
        _fPrev := _fLast; // 旧末帧降为前帧 / the old last to the previous
        _fLast := fIn; // 新样本入末帧 / the new sample to the last
        _bHave := TRUE; // 双帧齐备（第二帧起成立）/ the two samples ready
    ELSE // 非有限样本拒收（环不写、置位、计数，本库纪律②）/ a non finite sample rejected
        bBad := TRUE; // 置拒收实时标志 / raise the rejection flag
        IF nSkipCnt < DL_DRS_CNTMAX THEN // 计数防回绕 / the wrap guard
            nSkipCnt := nSkipCnt + 1; // 拒收计数推进 / advance the skip count
        END_IF
    END_IF
END_IF

// 段 4｜插值桥接输出（相位单点回夹 + 有限性闸，边界一二）/ segment 4, the interpolated bridge outlet
IF bEnable AND _bHave AND _bFin AND (_fPrev = _fPrev) AND ((_fPrev - _fPrev) = (_fPrev - _fPrev)) THEN // 双帧齐且有限 / both ready and finite
    IF fFrac < 0.0 THEN // 相位下越域回夹 / the phase below the band
        fFrac := 0.0; // 夹到零 / clamp to zero
        bClamped := TRUE; // 信息级 / informational
    ELSIF fFrac > 1.0 THEN // 相位上越域回夹 / the phase above the band
        fFrac := 1.0; // 夹到一 / clamp to one
        bClamped := TRUE; // 信息级 / informational
    END_IF
    fOut := _fPrev + (fFrac * (_fLast - _fPrev)); // 线性插值桥（不外推）/ the linear bridge, no extrapolation
    bValid := TRUE; // 输出可用 / the output usable
ELSE // 样本不足或非有限或失能：安全侧零 / not enough, non finite or disabled, the safe zero
    fOut := 0.0; // 安全侧零 / the safe zero
    bValid := FALSE; // 可用标志假 / the valid false
END_IF
END_FUNCTION_BLOCK

(* ---- FB_DL_DitherSignalGen.st ---- *)
// FB_DL_DitherSignalGen v1.0.0
// 开源溯源：self-cleanroom / 信号发生族补口
(*
  道莅工业代码库 | DL_MathData | FB_DL_DitherSignalGen
  版本: 1.0.0 | 日期: 2026-11-23 | 轮次: R75
  功能: 抖动信号发生（幅值/更新带宽可设）：LCG 伪随机数经更新节拍刷新，
        输出 ±幅值内均匀抖动，防 ADC 死区与摩擦滞环（dither 配套）
  邻件关系: 信号发生族 SineGenerator / PulseGenerator（确定性周期信号）——
            差异点：本件为伪随机幅值（LCG 32 位递推），非周期波形；
            更新带宽 = 更新节拍周期（1/ton 自复位周期）
  随机性声明: LCG 常数 a=1664525、c=1013904223（Numerical Recipes 公开口径），
            种子零值时自动注入非零初值防全零死锁
*)
FUNCTION_BLOCK FB_DL_DitherSignalGen
VAR_INPUT
    bEnable     : BOOL := FALSE;             // 使能（FALSE 输出回零）/ Enable, output to zero when FALSE
    fAmplitude  : REAL := 1.0;               // 抖动幅值 [工程单位]，域 > 0 / Dither amplitude, domain > 0
    tUpdate     : TIME := T#100MS;           // 更新节拍周期 [ms]，域 > 0 / Update tick period
    uSeed       : UDINT := 16#DEAD_BEEF;     // LCG 种子 [1]，0 时自动注入 / LCG seed, auto-inject when zero
END_VAR
VAR_OUTPUT
    fDitherOut  : REAL;                      // 抖动输出 ∈ [-幅值, +幅值] [工程单位] / Dither output within ±amplitude
    fNormRand   : REAL;                      // 归一随机数 ∈ [0,1] 诊断口 / Normalized random in [0,1]
    bTick       : BOOL;                      // 更新节拍脉冲（当拍到时单拍）/ Update tick pulse, one cycle
    bValid      : BOOL;                      // 组态有效回执 [-] / Config validity receipt
    bError      : BOOL;                      // 故障标志（组态非法）/ Fault flag (invalid config)
    uErrorId    : UDINT;                     // 事件码，0 = 无事件；16#0002_1F01 = 组态非法 / Event code
END_VAR
VAR
    uState      : UDINT;                     // LCG 当前状态 [1] / LCG current state
    bSeeded     : BOOL;                      // 已注入种子标志 [-] / Seeded flag
    tonTick     : TON;                       // 更新节拍定时器（自复位）/ Update tick timer, self-resetting
    fU          : REAL;                      // 归一随机中间量 [1] / Normalized random intermediate
END_VAR
VAR CONSTANT
    DL_DIT_LCG_A : UDINT := 16#0019_660D;    // LCG 乘数 a=1664525 [1] / LCG multiplier
    DL_DIT_LCG_C : UDINT := 16#3C6E_F35F;    // LCG 增量 c=1013904223 [1] / LCG increment
    DL_DIT_SCALE : REAL := 4294967295.0;     // 2^32-1 归一化分母 [1] / Normalization denominator
END_VAR

// —— 段 0：实例无条件刷新（R7：TON 每周期调用，IN := NOT Q 自复位） —— //
tonTick(IN := NOT tonTick.Q, PT := tUpdate);     // 节拍自复位（到时翻转一拍）/ Self-resetting tick timer
bTick := tonTick.Q;                              // 节拍脉冲单拍暴露 / Tick pulse exposed one cycle

// —— 段 1：组态闸 —— //
bValid := (fAmplitude > 0.0) AND (tUpdate > T#0MS) AND (fAmplitude = fAmplitude);   // 幅值正数 + 周期非零 + NaN 闸 / Gate
IF NOT bValid THEN
    bError   := TRUE;                            // 故障级：组态非法 / Fault level: invalid config
    uErrorId := 16#0002_1F01;                    // 故障码（1Fxx 步进）/ Fault code
    fDitherOut := 0.0;                           // 故障侧输出回零（安全位）/ Safe zero output
    fNormRand := 0.0;                            // 诊断口回零 / Diagnostic zero
    RETURN;
END_IF
bError   := FALSE;                               // 组态恢复：故障清零（解除路径）/ Fault cleared on valid config
uErrorId := 16#0000;                             // 事件码清零 / Event code cleared

// —— 段 2：种子注入（首拍或种子零值防死锁） —— //
IF (NOT bSeeded) OR (uState = 16#0000_0000) THEN
    IF uSeed = 16#0000_0000 THEN
        uState := 16#DEAD_BEEF;                  // 种子零值注入非零初值 / Inject nonzero on zero seed
    ELSE
        uState := uSeed;                         // 用户种子 / User seed
    END_IF
    bSeeded := TRUE;                             // 已注入标志 / Seeded flag
END_IF

// —— 段 3：使能与节拍驱动（节拍到时才刷新随机数，带宽即 1/tUpdate） —— //
IF NOT bEnable THEN
    fDitherOut := 0.0;                           // 失能输出回零（安全位）/ Disabled safe zero
    fNormRand := 0.0;                            // 诊断口回零 / Diagnostic zero
    RETURN;
END_IF
IF tonTick.Q THEN                                // 仅节拍拍刷新（拍间保持）/ Refresh only on tick, hold between
    uState := (uState * DL_DIT_LCG_A) + DL_DIT_LCG_C;    // LCG 递推（32 位自然回绕）/ LCG step, natural wrap
    fU := DWORD_TO_REAL(uState) / DL_DIT_SCALE;  // 归一化 ∈ [0,1] / Normalize to [0,1]
    IF fU > 1.0 THEN
        fU := 1.0;                               // 上钳（舍入防御）/ Clamp high
    END_IF
    fNormRand := fU;                             // 归一随机诊断口 / Diagnostic normalized random
    fDitherOut := (2.0 * fU - 1.0) * fAmplitude; // 映射 ±幅值（均匀分布）/ Map to ±amplitude uniform
END_IF
END_FUNCTION_BLOCK

(* ---- FB_DL_EventRateCalc.st ---- *)
(*==============================================================================
 * 组件名称 (Component)  : FB_DL_EventRateCalc
 * 溯源说明 (Provenance) : IEC 61131-3 标准语义的道莅防御性实现（零检索变体线）
 * 所属子库 (Sublibrary) : DL_MathData / Statistics
 * 当前版本 (Version)    : 1.0.0
 * 兼容性   (Platform)   : CODESYS 3.5 / TwinCAT 3 / 汇川 InoProShop；
 *                         纯 IEC 61131-3（第 3 版），仅用标准库 TON / R_TRIG
 * 组件分类 (Category)   : 功能块（FUNCTION_BLOCK）· 滑窗事件速率
 * 功能一句话 (Summary)  : 环形 60 桶滑窗事件计数，输出事件每分钟速率与累计数。
 * 边界与安全 (Boundary) : ①窗口小于 1 s 钳 1 s；大于 1 h 钳 1 h，均置钳位码；
 *                         ②钳位后继续正常工作（码级不断链）；
 *                         ③bReset 清全部桶、速率与累计；
 *                         ④桶推进定时器与事件沿检测均无条件周期刷新；
 *                         ⑤窗口时长为 0 防御（除零前判）。
 * 错误码    : 16#0001_03C3 窗口钳位发生（1 s 或 1 h 边界）——故障级（持续态）
 *             16#0001_03C4 保留禁用（不得挪用，本件零赋值）
 * 码位总账  : 16#0001_03C3 用 ｜ 16#0001_03C4 预留
 * 修改记录  : v1.0.0 R26 初版
 *==============================================================================*)
FUNCTION_BLOCK FB_DL_EventRateCalc
VAR_INPUT
    bEvent  : BOOL;   // 事件脉冲输入（内部取上升沿）/ Event pulse input (edge taken inside)
    tWindow : TIME;   // 滑窗时长 1 s~1 h，越界钳位 [ms] / Sliding window 1 s to 1 h, clamped
    bReset  : BOOL;   // 复位：清桶、速率与累计 / Reset: clear buckets, rate and total
END_VAR
VAR_OUTPUT
    fRate  : LREAL; // 事件速率（事件每分钟）/ Event rate (events per minute)
    uTotal : ULINT; // 累计事件总数 / Total accumulated events
    eErr   : UDINT; // 本周期错误码，0=无错 / Error code this cycle, 0 = none
END_VAR
VAR CONSTANT
    cBuckets   : INT := 60;        // 环形桶数（固定）/ Fixed ring bucket count
    cMsMin     : DINT := 1000;     // 窗口下限 1 s [ms] / Window lower bound 1 s [ms]
    cMsMax     : DINT := 3600000;  // 窗口上限 1 h [ms] / Window upper bound 1 h [ms]
END_VAR
VAR
    aBuckets   : ARRAY[0..59] OF ULINT; // 环形计数桶 / Ring counting buckets
    iHead      : INT;            // 当前桶索引 / Current bucket index
    tonBkt     : TON;            // 桶推进定时器（无条件刷新）/ Bucket advance timer (unconditional refresh)
    rTrigEvt   : R_TRIG;         // 事件上升沿检测（无条件刷新）/ Event rising edge (unconditional refresh)
    dwWinMs    : DINT;           // 窗口有效时长 [ms] / Effective window duration [ms]
    dwBktMs    : DINT;           // 单桶时长 [ms] / Per-bucket duration [ms]
    i          : INT;            // 求和游标 / Summation cursor
    uSum       : ULINT;          // 窗口内事件合计 / Events summed over window
    fWinSec    : LREAL;          // 窗口时长秒值（速率换算分母）/ Window seconds (rate denominator)
END_VAR

// ---------- 无条件周期刷新：沿检测 + 桶推进定时器 ----------
rTrigEvt(CLK := bEvent);
dwWinMs := TIME_TO_DINT(tWindow);            // 窗口毫秒读数 / Window in milliseconds

// ---------- 窗口钳位防御（先钳后用，码级持续态） ----------
eErr := 0;
IF dwWinMs < cMsMin THEN
    dwWinMs := cMsMin;                       // 下限钳 1 s / Clamp to 1 s lower bound
    eErr    := 16#0001_03C3;                 // 钳位码 / Clamp code
ELSIF dwWinMs > cMsMax THEN
    dwWinMs := cMsMax;                       // 上限钳 1 h / Clamp to 1 h upper bound
    eErr    := 16#0001_03C3;                 // 钳位码（复用同码）/ Clamp code (shared)
END_IF

// ---------- 复位优先：清桶清累计清速率 ----------
IF bReset THEN
    FOR i := 0 TO cBuckets - 1 DO
        aBuckets[i] := 0;                    // 清所有桶 / Clear all buckets
    END_FOR
    iHead  := 0;                             // 桶头归零 / Head index reset
    uTotal := 0;                             // 累计清零 / Total cleared
    fRate  := 0.0;                           // 速率清零 / Rate cleared
END_IF

// ---------- 桶推进：单桶时长 = 窗口 / 桶数（除零前判） ----------
IF dwWinMs > 0 THEN
    dwBktMs := dwWinMs / cBuckets;           // 整除单桶毫秒 / Integer per-bucket ms
ELSE
    dwBktMs := cMsMin;                       // 防御缺省（理论不可达）/ Defensive default
END_IF
tonBkt(IN := TRUE, PT := DINT_TO_TIME(dwBktMs));
IF tonBkt.Q THEN
    iHead := (iHead + 1) MOD cBuckets;       // 环形推进 / Ring advance
    aBuckets[iHead] := 0;                    // 新桶清零（旧桶自然滑出窗）/ New bucket cleared
END_IF

// ---------- 事件入桶：沿触发计数，累计同步递增 ----------
IF rTrigEvt.Q THEN
    aBuckets[iHead] := aBuckets[iHead] + 1;  // 当前桶计数加一 / Increment current bucket
    uTotal := uTotal + 1;                    // 累计事件加一 / Total incremented
END_IF

// ---------- 速率换算：窗口合计 / 窗口分钟数（分母前判零） ----------
uSum := 0;
FOR i := 0 TO cBuckets - 1 DO
    uSum := uSum + aBuckets[i];              // 窗口合计 / Window sum
END_FOR
fWinSec := ULINT_TO_LREAL(DINT_TO_ULINT(dwWinMs)) / 1000.0; // 窗口秒值 / Window seconds
IF fWinSec > 0.0 THEN
    fRate := ULINT_TO_LREAL(uSum) * 60.0 / fWinSec;    // 事件每分钟 / Events per minute
ELSE
    fRate := 0.0;                            // 除零防御缺省 / Divide-by-zero guard default
END_IF

END_FUNCTION_BLOCK

(* ---- FB_DL_FirstOrderImpResp.st ---- *)
// FB_DL_FirstOrderImpResp v1.0.0
// 开源溯源：brOscatLib / URL https://github.com/iec-oscat-mirror / 许可证 MIT / 借鉴 FT_IMP 一阶惯性环节脉冲响应语义，clean-room 重写
(*
  道莅工业代码库 | DL_MathData | FB_DL_FirstOrderImpResp
  版本: 1.0.0 | 日期: 2026-11-23 | 轮次: R75
  功能: 一阶惯性环节脉冲响应序列计算：h(t) = (K/T)·e^(-t/T)，采样 t_k = k·Ts
  邻件关系: 与 FB_DL_FirstOrderIdent 同族不同用 —— 辨识件由数据反推 K/T，
            本件由 K/T 正推响应序列（辨识 vs 响应），口径互不引用
  接口契约: bExecute 上升沿触发整段序列计算（单拍完成，非逐拍递推）；
            nLen 为本次计算点数，域 1..64，超域按 64 钳位并置信息码
*)
FUNCTION_BLOCK FB_DL_FirstOrderImpResp
VAR_INPUT
    bExecute  : BOOL := FALSE;                   // 执行触发（上升沿整段计算）/ Execute trigger, rising edge
    fGain     : REAL := 1.0;                     // 增益 K [1]，域 > 0 / DC gain, domain > 0
    fTimeConst: REAL := 1.0;                     // 时间常数 T [s]，域 > 0 / Time constant [s]
    fTs       : REAL := 0.1;                     // 采样周期 Ts [s]，域 > 0 / Sampling period [s]
    nLen      : INT := 16;                       // 序列点数 [点]，域 1..64 / Sequence length [points], domain 1..64
END_VAR
VAR_OUTPUT
    aResp     : ARRAY[1..64] OF REAL;            // 脉冲响应序列 h(t_k) [1/s·(s/点)，随增益] / Impulse response sequence
    nCount    : INT;                             // 本次实际写出点数 [点] / Actual points written
    bDone     : BOOL;                            // 本次序列计算完成脉冲（单拍自清）/ Sequence done pulse, one cycle
    bValid    : BOOL;                            // 参数有效且序列可用 [-] / Parameters valid and sequence usable
    bError    : BOOL;                            // 故障标志，与故障级码配对 / Fault flag paired with fault code
    uErrorId  : UDINT;                           // 事件码，0 = 无事件 / Event code, 0 = none
END_VAR
VAR
    rtrExec   : R_TRIG;                          // 执行沿检测（每拍无条件刷新）/ Execute edge, refreshed every cycle
    bCfgOk    : BOOL;                            // 参数闸结果 [-] / Parameter gate result
    nLenEff   : INT;                             // 钳位后生效点数 [点] / Effective clamped length
    fDecay    : REAL;                            // 单步衰减因子 e^(-Ts/T) [1] / Per-step decay factor
    fPeak     : REAL;                            // 脉冲响应峰值 K/T [1/s] / Impulse peak K/T
    fTerm     : REAL;                            // 当前项 K/T·decay^k [1/s] / Current term
    i         : INT;                             // 循环索引 [点] / Loop index
END_VAR
VAR CONSTANT
    DL_FIR_LENMAX : INT := 64;                   // 序列上限（数组显式上界一致）[点] / Sequence upper bound, matches array
END_VAR

// —— 段 0：实例无条件刷新 + 输出缺省 —— //
rtrExec(CLK := bExecute);                        // 执行沿每拍刷新 / Execute edge refreshed every cycle
bDone := FALSE;                                  // 完成脉冲单拍自清 / Done pulse self-clearing

// —— 段 1：参数闸（有限性 + 正数域 + 点数域） —— //
bCfgOk := (fGain > 0.0) AND (fTimeConst > 0.0) AND (fTs > 0.0)
          AND (fGain = fGain) AND (fTimeConst = fTimeConst) AND (fTs = fTs);   // 正数域 + NaN 自反判 / Positive domain and NaN gate
bValid := bCfgOk;                                // 有效回执随参数闸 / Validity follows gate
IF NOT bCfgOk THEN
    bError   := TRUE;                            // 故障级：参数非法 / Fault level: invalid parameters
    uErrorId := 16#0002_1A01;                    // 本件故障码（1Axx 步进）/ Fault code of this component
    RETURN;                                      // 参数非法不计算 / No calculation on invalid params
END_IF
bError   := FALSE;                               // 参数恢复：故障清零（解除路径）/ Fault cleared on valid params
uErrorId := 16#0000;                             // 事件码清零 / Event code cleared
nLenEff := nLen;                                 // 生效点数初值 / Effective length init
IF nLenEff < 1 THEN
    nLenEff := 1;                                // 下限钳位 / Clamp to lower bound
END_IF
IF nLenEff > DL_FIR_LENMAX THEN
    nLenEff := DL_FIR_LENMAX;                    // 上限钳位至数组上界 / Clamp to array bound
END_IF
nCount := nLenEff;                               // 实际点数输出 / Actual count output

// —— 段 2：上升沿触发整段序列计算 —— //
IF rtrExec.Q THEN                                // 仅执行沿拍计算（避免每拍重算）/ Compute only on execute edge
    fDecay := EXP(-fTs / fTimeConst);            // 单步衰减 e^(-Ts/T)，T 非零已过闸 / Per-step decay, T nonzero gated
    fPeak  := fGain / fTimeConst;                // 峰值 K/T / Peak value K/T
    fTerm  := fPeak;                             // 首项 k=0 / First term k=0
    FOR i := 1 TO nLenEff DO                       // 逐点写出（显式上界，无 VLA）/ Write points with explicit bound
        aResp[i] := fTerm;                       // h(t_k) = (K/T)·e^(-k·Ts/T) / Sampled impulse response
        fTerm := fTerm * fDecay;                 // 迭代衰减（避免逐点 EXP 开销）/ Iterative decay
    END_FOR
    bDone := TRUE;                               // 完成脉冲（单拍，段 0 下拍自清）/ Done pulse for one cycle
END_IF
END_FUNCTION_BLOCK

(* ---- FB_DL_HistogramAccum.st ---- *)
(*==============================================================================
 * 组件名称 (Component)  : FB_DL_HistogramAccum
 * 溯源说明 (Provenance) : 道莅 clean-room 防御性实现（LGF Measurement 统计族深化）
 * 所属子库 (Sublibrary) : DL_MathData / Statistics
 * 当前版本 (Version)    : 1.0.0
 * 兼容性   (Platform)   : CODESYS 3.5 / TwinCAT 3 / 汇川 InoProShop；
 *                         纯 IEC 61131-3（第 3 版），零标准库依赖
 * 组件分类 (Category)   : 功能块（FUNCTION_BLOCK）· 数值直方图累积
 * 功能一句话 (Summary)  : 按单调递增边界表分箱加权计数，含下溢/上溢桶与非有限拦截。
 * 边界与安全 (Boundary) : ①NaN 拒收（x <> x 自反判）与无穷拒收（差值自反判）；
 *                         ②权重非正拒收（复用样本非法码，R90 口径）；
 *                         ③边界表未单调递增 → bEdgeErr 且本拍不累计；
 *                         ④右闭约定：值恰等于边界归上侧箱（右箱）；
 *                         ⑤数组下标全程钳位，禁越界写；
 *                         ⑥容量上限 64 箱，超容箱计入上溢。
 * 错误码    : 16#0001_03C5 样本拒收（NaN/无穷/权重非正）——故障级（持续态）
 *             16#0001_03C6 边界表非法（未单调递增或点数不足）——故障级（持续态）
 * 码位总账  : 16#0001_03C5 用 ｜ 16#0001_03C6 用
 * 修改记录  : v1.0.0 R26 初版
 *==============================================================================*)
FUNCTION_BLOCK FB_DL_HistogramAccum
VAR_INPUT
    fValue  : LREAL;  // 待分箱样本值 / Sample value to bin
    fWeight : LREAL;  // 样本权重，默认 1.0 / Sample weight, default 1.0
    bReset  : BOOL;   // 复位：清全部计数 / Reset: clear all counts
END_VAR
VAR_IN_OUT
    aEdges  : ARRAY[*] OF LREAL; // 单调递增分箱边界表 / Monotonic increasing bin edges
END_VAR
VAR_OUTPUT
    aCounts    : ARRAY[*] OF ULINT; // 各箱计数（与边界表同界）/ Counts per bin (same bounds as edges)
    uUnderflow : ULINT; // 下溢桶：低于最小边界的计数 / Underflow bucket count
    uOverflow  : ULINT; // 上溢桶：高于最大边界的计数 / Overflow bucket count
    bEdgeErr   : BOOL;  // 边界表非法标志（未单调递增）/ Illegal edge table flag
    eErr       : UDINT; // 本周期错误码，0=无错 / Error code this cycle, 0 = none
END_VAR
VAR CONSTANT
    cMaxBins : INT := 64; // 内部容量上限 64 箱 / Internal capacity limit 64 bins
END_VAR
VAR
    aCntBuf   : ARRAY[0..63] OF ULINT; // 内部计数缓冲（跨拍保持）/ Internal counts buffer (kept across scans)
    uUfBuf    : ULINT; // 内部下溢计数 / Internal underflow count
    uOfBuf    : ULINT; // 内部上溢计数 / Internal overflow count
    nEdges    : INT;   // 边界点数 / Edge point count
    i         : INT;   // 分箱搜索游标 / Bin search cursor
    iUb       : INT;   // 输出数组上界 / Output array upper bound
    bSorted   : BOOL;  // 边界单调性中间判据 / Edge monotonicity intermediate
    bAccumOk  : BOOL;  // 本拍允许累计判据 / Accumulation allowed this cycle
END_VAR

// ---------- 周期起点：错误码与标志先清（持续态随后重置） ----------
eErr     := 0;
bEdgeErr := FALSE;
bAccumOk := TRUE;

// ---------- 复位优先：清内部计数 ----------
IF bReset THEN
    FOR i := 0 TO cMaxBins - 1 DO
        aCntBuf[i] := 0;                     // 清内部箱 / Clear internal bins
    END_FOR
    uUfBuf := 0;                             // 清下溢 / Clear underflow
    uOfBuf := 0;                             // 清上溢 / Clear overflow
END_IF

// ---------- 边界表防御：点数与单调性（下标钳位访问） ----------
nEdges := UPPER_BOUND(aEdges, 1) + 1;        // 边界点数 / Edge point count
IF nEdges < 2 THEN
    bEdgeErr := TRUE;                        // 点数不足 / Insufficient points
    eErr     := 16#0001_03C6;                // 边界表非法 / Illegal edge table
ELSE
    bSorted := TRUE;
    FOR i := 0 TO nEdges - 2 DO
        IF NOT (aEdges[i] < aEdges[i + 1]) THEN
            bSorted := FALSE;                // 严格递增被破坏 / Strict increase violated
        END_IF
    END_FOR
    IF NOT bSorted THEN
        bEdgeErr := TRUE;                    // 置非法标志 / Set illegal flag
        eErr     := 16#0001_03C6;            // 边界表非法码 / Illegal table code
    END_IF
END_IF
IF bEdgeErr THEN
    bAccumOk := FALSE;                       // 表非法本拍不累计 / No accumulation on illegal table
END_IF

// ---------- 样本防御：非有限与权重（拒收不累计） ----------
IF bAccumOk THEN
    IF (fValue <> fValue) OR ((fValue - fValue) <> (fValue - fValue)) THEN
        bAccumOk := FALSE;                   // NaN 或无穷拒收 / NaN or Inf rejected
        eErr     := 16#0001_03C5;            // 样本非法码 / Illegal sample code
    ELSIF (fWeight <= 0.0) OR (fWeight <> fWeight) THEN
        bAccumOk := FALSE;                   // 权重非正拒收（复用 03C5）/ Non-positive weight rejected (03C5 reuse)
        eErr     := 16#0001_03C5;            // 样本非法码（R90 复用）/ Illegal sample code (R90 reuse)
    END_IF
END_IF

// ---------- 分箱累计：右闭约定，恰等边界归右箱 ----------
IF bAccumOk THEN
    IF fValue < aEdges[0] THEN
        uUfBuf := uUfBuf + ULINT#1; // 低于最小边界 → 下溢 / Below first edge: underflow
    ELSIF fValue > aEdges[nEdges - 1] THEN
        uOfBuf := uOfBuf + ULINT#1; // 高于最大边界 → 上溢 / Above last edge: overflow
    ELSE
        i := 0;
        WHILE (i < nEdges - 1) AND (fValue > aEdges[i]) DO
            i := i + 1;                      // 找首个上边界不小于值的箱 / Find first upper edge covering value
        END_WHILE
        IF i > cMaxBins - 1 THEN
            i := cMaxBins - 1;               // 下标钳位，超容归上溢侧 / Clamp index, over-capacity to overflow
            uOfBuf := uOfBuf + ULINT#1;
        ELSE
            aCntBuf[i] := aCntBuf[i] + LREAL_TO_ULINT(fWeight); // 加权计数 / Weighted count
        END_IF
    END_IF
END_IF

// ---------- 输出镜像：按输出数组实际界钳位拷贝 ----------
iUb := UPPER_BOUND(aCounts, 1);
IF iUb > cMaxBins - 1 THEN
    iUb := cMaxBins - 1;                     // 输出上界钳位 / Clamp output upper bound
END_IF
FOR i := 0 TO iUb DO
    aCounts[i] := aCntBuf[i];                // 内部缓冲镜像到输出 / Mirror buffer to outputs
END_FOR
uUnderflow := uUfBuf;                        // 下溢输出 / Underflow output
uOverflow  := uOfBuf;                        // 上溢输出 / Overflow output

END_FUNCTION_BLOCK

(* ---- FB_DL_HistogramBinTally.st ---- *)
(*
  Name        : FB_DL_HistogramBinTally
  Category    : DL_MathData
  Version     : 1.0.0
  Purpose     : 分箱直方图累计：等宽 bins 样本逐拍落格计数，越界钳边计数，占比出口按总入格数派生；/ Histogram bin tally: equal-width bins with per-scan sample counting, clamped-edge counting, and ratio outlets derived from total tally
  溯源        : 借 lgf-measurement 的统计族扩组织，clean-room 实现
  Boundary    : ① bins 数域 2..64 且 bin 宽 > 0，任一越域锁存故障（计数值冻结不动）；
                ② 落格下标由边界值直比算出（FOR 逐格上界直比，不用除法），越下界钳第 1 格、越上界钳末格，同时钳边计数出口分别累加；
                ③ 非有限样本拒收不入格（bSampleRej 单拍脉冲，R187 出口映射）；
                ④ 复位沿幂等清零：计数出口与内部计数器同拍同步归零（防镜像失步）；
                ⑤ 占比除子 = 总入格数，总数 0 时占比出口全 0 不除（防除零）；
                ⑥ 计数器为 UDINT 饱和累加（达上限不再递增，防回卷）。
*)
TYPE E_DL_HbtState :
(
    eIdle  := 0,                             (* 未使能（计数清零保持） / Disabled, tallies cleared *)
    eRun   := 10,                            (* 直方图累计运行 / Tally running *)
    eFault := 90                             (* 故障锁存相 / Fault latched *)
);
END_TYPE

TYPE E_DL_HbtCause :
(
    eNone      := 0,                         (* 无故障成因 / No cause *)
    eCfgIllegal:= 1,                        (* 组态非法：bins/格宽越域 / Illegal config *)
    ePhaseBad  := 2                         (* 非法相位兜底 / Illegal phase fallback *)
);
END_TYPE

FUNCTION_BLOCK FB_DL_HistogramBinTally
VAR_INPUT
    fSample : REAL := 0.0;                   (* 样本输入（任意工程量）[-] / Sample input *)
    fLower  : REAL := 0.0;                   (* 第 1 格下边界 [工程单位] / Lower edge of bin 1 *)
    fBinW   : REAL := 1.0;                   (* 等宽格宽，域 > 0 [工程单位] / Bin width *)
    nBins   : INT := 16;                     (* 格数，域 2..64 [格] / Bin count *)
    bEnable : BOOL := TRUE;                  (* 使能 [-] / Enable *)
    bReset  : BOOL := FALSE;                 (* 复位命令，上升沿幂等清零 [-] / Reset command *)
END_VAR
VAR_OUTPUT
    aBinCnt : ARRAY[1..64] OF UDINT;         (* 各格计数（有效区 1..nBins，其余恒 0）[个] / Bin tallies *)
    nTotal  : UDINT;                         (* 总入格数（含钳边，不含拒收）[个] / Total tallied count *)
    nClampLow: UDINT;                        (* 越下界钳第 1 格累计数 [个] / Clamped-low count *)
    nClampHigh: UDINT;                       (* 越上界钳末格累计数 [个] / Clamped-high count *)
    nLastBin: INT;                           (* 最近样本落格序号（0 = 拒收/未落格）[格] / Last sample bin index *)
    fLastRatio: REAL;                        (* 最近落格占比 = 该格计数 / 总入格数 [-] / Last bin ratio *)
    bSampleRej: BOOL;                        (* 最近样本被拒收（单拍脉冲）[-] / Sample rejected pulse *)
    eState  : E_DL_HbtState;                 (* 状态出口 / State outlet *)
    eCause  : E_DL_HbtCause;                 (* 故障成因出口（R190 归因唯一） / Fault cause outlet *)
    bError  : BOOL;                          (* 故障锁存标志 [-] / Fault latch flag *)
END_VAR
VAR
    _eState : E_DL_HbtState := E_DL_HbtState.eIdle;  (* 内部相位（CASE 唯一写入目标） / Internal phase *)
    _eCause : E_DL_HbtCause := E_DL_HbtCause.eNone;  (* 故障成因锁存量 / Latched cause *)
    rtReset : R_TRIG;                        (* 复位沿实例，段 0 无条件调用 / Reset edge instance *)
    _bFault : BOOL;                          (* 故障锁存位 / Latched fault bit *)
    _bCfgBad: BOOL;                          (* 组态非法当拍量 / Illegal config this scan *)
    _bFin   : BOOL;                          (* 样本有限性当拍量 / Sample finiteness *)
    _bRejI  : BOOL;                          (* 拒收脉冲内部量（统一出口映射，R187） / Reject pulse internal *)
    _bHit   : BOOL;                          (* 本拍落格成功当拍量 / Binned this scan *)
    _nBin   : INT;                           (* 本拍落格序号 [格] / Bin index this scan *)
    _i      : INT;                           (* 落格扫描游标 [格] / Bin scan cursor *)
    _nBinsE : INT;                           (* 钳位后生效格数 [格] / Effective bin count *)
    _nCntI  : UDINT;                         (* 落格计数中间量（占比派生用）[个] / Bin count intermediate *)
END_VAR
VAR CONSTANT
    DL_HBT_NMIN : INT   := 2;                (* 格数下限（边界①）[格] / Bin count lower bound *)
    DL_HBT_NMAX : INT   := 64;               (* 格数上限（边界①）[格] / Bin count upper bound *)
    DL_HBT_EPS  : REAL  := 1.0E-6;           (* 判零容差 [-] / Epsilon *)
    DL_HBT_CNTMAX: UDINT := 4294967295;      (* 计数饱和上限（边界⑥，R28）[个] / Tally saturation cap *)
END_VAR

(* —— 段 0：当拍判据派生 + 实例无条件刷新（R228A） —— *)
_bCfgBad := (nBins < DL_HBT_NMIN) OR (nBins > DL_HBT_NMAX) OR (fBinW <= DL_HBT_EPS);   (* 格数/格宽域闸（边界①） / Bin count and width gates *)
rtReset(CLK := bReset);                                  (* 复位沿每拍必调 / Reset edge every scan *)
_bFin := (fSample = fSample) AND ((fSample - fSample) = (fSample - fSample));   (* 样本 NaN 自反 + Inf 差判闸（边界③） / Sample NaN and Inf gate *)
_nBinsE := nBins;                                        (* 生效格数初值 / Effective bins init *)
IF _nBinsE < DL_HBT_NMIN THEN
    _nBinsE := DL_HBT_NMIN;                              (* 格数下限钳位（防越界） / Bin count lower clamp *)
END_IF
IF _nBinsE > DL_HBT_NMAX THEN
    _nBinsE := DL_HBT_NMAX;                              (* 格数上限钳位（防越界） / Bin count upper clamp *)
END_IF

(* —— 段 1：单拍量预清零（R107） —— *)
_bRejI := FALSE;                                         (* 拒收脉冲内部量预清 / Reject pulse preset *)
bSampleRej := FALSE;                                     (* 拒收脉冲出口预清 / Reject outlet preset *)
nLastBin := 0;                                           (* 落格序号预清（拒收拍为 0） / Bin index preset *)
fLastRatio := 0.0;                                       (* 占比出口预清（除子零保护默认） / Ratio preset zero *)
_bHit := FALSE;                                          (* 落格成功量预清 / Binned preset *)
_nBin := 0;                                              (* 落格序号中间量预清 / Bin index intermediate *)

(* —— 段 2：复位沿处理（作用域：清故障 + 全计数出口与内部同拍归零，R283/边界④） —— *)
IF rtReset.Q THEN
    _bFault := FALSE;                                    (* 清故障锁存 / Clear fault *)
    _eCause := E_DL_HbtCause.eNone;                      (* 清成因 / Clear cause *)
    FOR _i := 1 TO DL_HBT_NMAX DO
        aBinCnt[_i] := UDINT#0;                          (* 各格计数同拍归零（幂等） / Bin tallies zeroed *)
    END_FOR
    nTotal := UDINT#0;                                   (* 总入格数归零 / Total zeroed *)
    nClampLow := UDINT#0;                                (* 钳下界计数归零 / Clamp-low zeroed *)
    nClampHigh := UDINT#0;                               (* 钳上界计数归零 / Clamp-high zeroed *)
    nLastBin := 0;                                       (* 落格序号归零 / Bin index zeroed *)
    fLastRatio := 0.0;                                   (* 占比归零 / Ratio zeroed *)
    _eState := E_DL_HbtState.eIdle;                      (* 迁未使能相 / Back to idle *)
END_IF

(* —— 段 3：组态故障锁存（锁存至复位沿，R189） —— *)
IF _bCfgBad AND NOT _bFault THEN
    _bFault := TRUE;                                     (* 锁存故障位 / Latch fault *)
    _eCause := E_DL_HbtCause.eCfgIllegal;                (* 成因：组态非法 / Cause illegal config *)
    _eState := E_DL_HbtState.eFault;                     (* 同步迁故障相 / Migrate to fault *)
END_IF

(* —— 段 4：CASE 主状态机（ELSE 兜底迁 eFault，红线 6） —— *)
CASE _eState OF
    E_DL_HbtState.eIdle:                                 (* 未使能：计数清零保持（不留陈旧） / Disabled *)
        FOR _i := 1 TO DL_HBT_NMAX DO
            aBinCnt[_i] := UDINT#0;                      (* 失能各格计数清零 / Disabled tallies cleared *)
        END_FOR
        nTotal := UDINT#0;                               (* 失能总数清零 / Disabled total cleared *)
        nClampLow := UDINT#0;                            (* 失能钳下界清零 / Disabled clamp-low cleared *)
        nClampHigh := UDINT#0;                           (* 失能钳上界清零 / Disabled clamp-high cleared *)
        IF bEnable AND NOT _bFault THEN
            _eState := E_DL_HbtState.eRun;               (* 进入累计相 / Enter running *)
        END_IF
    E_DL_HbtState.eRun:                                  (* 累计相：逐拍落格 / Running *)
        IF NOT bEnable THEN
            _eState := E_DL_HbtState.eIdle;              (* 失能回未使能 / Back to idle *)
        ELSIF _bFin THEN                                 (* 非有限样本整拍拒收（边界③） / Non-finite rejected *)
            FOR _i := 1 TO _nBinsE DO                    (* 边界值直比找格（不用除法，边界②） / Edge compare binning *)
                IF fSample < (fLower + fBinW * INT_TO_REAL(_i)) THEN
                    _nBin := _i;                         (* 首个上界大于样本的格即落格 / First upper edge above sample *)
                    _bHit := TRUE;                       (* 落格成功 / Binned *)
                    EXIT;
                END_IF
            END_FOR
            IF NOT _bHit THEN
                IF fSample < fLower THEN
                    _nBin := 1;                          (* 越下界钳第 1 格（边界②） / Clamp to bin 1 *)
                    IF nClampLow < DL_HBT_CNTMAX THEN
                        nClampLow := nClampLow + UDINT#1;    (* 钳下界计数饱和累加 / Clamp-low tally *)
                    END_IF
                ELSE
                    _nBin := _nBinsE;                    (* 越上界钳末格（边界②） / Clamp to last bin *)
                    IF nClampHigh < DL_HBT_CNTMAX THEN
                        nClampHigh := nClampHigh + UDINT#1;  (* 钳上界计数饱和累加 / Clamp-high tally *)
                    END_IF
                END_IF
                _bHit := TRUE;                           (* 钳边落格成功 / Clamped binned *)
            END_IF
            IF _bHit AND (_nBin >= 1) AND (_nBin <= _nBinsE) THEN    (* 双重下标域闸（防越界写） / Index domain gate *)
                IF aBinCnt[_nBin] < DL_HBT_CNTMAX THEN
                    aBinCnt[_nBin] := aBinCnt[_nBin] + UDINT#1;      (* 该格计数饱和累加 / Bin tally *)
                END_IF
                IF nTotal < DL_HBT_CNTMAX THEN
                    nTotal := nTotal + UDINT#1;          (* 总入格数饱和累加 / Total tally *)
                END_IF
                nLastBin := _nBin;                       (* 落格序号出口 / Bin index outlet *)
                _nCntI := aBinCnt[_nBin];                (* 占比分子中间量 / Ratio numerator *)
                IF nTotal > UDINT#0 THEN                 (* 占比除子 = 总数，零保护（边界⑤） / Ratio divisor gate *)
                    fLastRatio := _nCntI / UDINT_TO_REAL(nTotal);    (* 占比派生（除子已过闸） / Ratio derived *)
                END_IF
            END_IF
        ELSE
            _bRejI := TRUE;                              (* 非有限拍置拒收内部脉冲（R187） / Reject internal pulse *)
        END_IF
    E_DL_HbtState.eFault:                                (* 故障相：计数冻结保持，仅复位沿出 / Fault *)
        ;                                                (* 锁存回放（R28） / Replay from latch *)
    ELSE                                                 (* 非法相位兜底迁安全态 / Illegal phase fallback *)
        _eState := E_DL_HbtState.eFault; _bFault := TRUE;    (* 迁故障相 + 同步锁存 / To fault and latch *)
        _eCause := E_DL_HbtCause.ePhaseBad;              (* 成因：非法相位 / Cause illegal phase *)
END_CASE

(* —— 段 5：出口映射（内部 _b* → 输出单拍，R187；名实双出口，R191） —— *)
bSampleRej := _bRejI;                                    (* 拒收脉冲单拍出口 / Reject pulse outlet *)
bError := _bFault;                                       (* 故障标志镜像 / Fault flag mirror *)
eState := _eState;                                       (* 状态出口 / State outlet *)
eCause := _eCause;                                       (* 成因出口 / Cause outlet *)
END_FUNCTION_BLOCK

(* ---- FB_DL_LifoStack.st ---- *)
(*==============================================================================
 * 组件名称 (Component)  : FB_DL_LifoStack
 * 所属子库 (Sublibrary) : DL_MathData
 * 当前版本 (Version)    : 1.0.0
 * 兼容性   (Platform)   : CODESYS 3.5 / TwinCAT 3 / 汇川 InoProShop / Machine Expert
 *                         仅依赖 Standard.library（R_TRIG），无厂商方言
 * 功能描述 (Function)   : 定长 64 深度 LIFO 栈（后进先出），支持压栈、弹栈、
 *                         窥视栈顶、清空四操作，全部 O(1)，无任何元素搬移。
 *                         带上溢/下溢锁存与单调累计计数。用于工艺路径回溯
 *                         （走了哪些工位、原路退回）、嵌套配方解析、报警确认
 *                         的"撤销"语义、深度优先搜索的待办表。
 *                         满栈压入拒绝且不覆盖栈底：LIFO 无"丢最旧"语义，
 *                         静默覆盖会让路径回溯错位一格，现场极难排查。
 * 本文件内含       : E_DL_StackState（枚举，归属本组件）
 *                    FB_DL_LifoStack（功能块主体）
 * 开源溯源 (Origin)     : 原创实现（参考西门子 LGF 数据处理组的 FIFO/LIFO
 *                         拆分方式与"满/空/长度"状态位粒度，clean-room 编写，
 *                         未复制任何源码）。
 * 依赖     (Depends)    : 无 DL_ 内部依赖；Standard.library: R_TRIG
 * 红线自检 (Redline)    : R1 ✓ 零全局变量表与外部变量引用 ｜ R2 ✓ 零物理 IO 地址直写
 *                         R3 ✓ 纯 IEC 61131-3，计数比较显式转换 ｜ R4 ✓ 下标双检 + 空满拒绝
 *                         R5 ✓ 全变量中英双语同行注释 ｜ R6 ✓ ENUM + CASE + ELSE 兜底
 *                         R7 ✓ 两 R_TRIG 主体最前部无条件刷新
 *
 * 【与 FIFO 的区别 / Difference to FIFO（边界 B7）】
 *   同一序列 1,2,3 依次压入：FIFO（FB_DL_RingBufferLReal）弹出 1,2,3；
 *   本块弹出 3,2,1。本块只有单栈顶指针、无回绕，读/写双指针结构见环形队列块。
 *
 * 【同周期压弹次序 / Push-before-pop ordering（边界 B3）】
 *   同一扫描周期同时出现压栈沿与弹栈沿时，先压后弹：弹出的是刚压入的值。
 *   这是"写入后立即读回校验"的常见用法；次序不可交换，先弹后压会读到
 *   旧栈顶，调用方会误判校验失败。
 *
 * 【哨兵值披露 / Sentinel disclosure（边界 B2）】
 *   空栈时栈顶输出 0.0、下溢弹出值输出 0.0，该 0.0 是哨兵不是数据。
 *   判空必须看空标志或深度计数，不得以"栈顶等于 0"反推栈状态。
 *
 * 【锁存纪律 / Latch discipline（边界 B5）】
 *   上溢/下溢故障码为锁存码，bClear 是唯一清锁存路径；清空保留
 *   累计计数（生命周期统计不清零）。
 * 修订历史 (Revision)   :
 *   2026-11-14  v1.0.0  首版入库（Phase 1 收口批次 · R3）
 *============================================================================*)
TYPE E_DL_StackState :
(
    eEmpty := 0,      // 空栈，无可弹数据 / Empty, nothing to pop
    eReady := 10,     // 有数据可弹 / Has data available
    eFault := 99      // 上溢或下溢锁存，需 bClear 解除 / Overflow or underflow latched, clear required
);
END_TYPE

FUNCTION_BLOCK FB_DL_LifoStack
VAR_INPUT
    bPush      : BOOL;                     // 上升沿：压入 fPushValue / Rising edge: push value
    fPushValue : LREAL := 0.0;             // 待压入值 [EU] / Value to push [EU]
    bPop       : BOOL;                     // 上升沿：弹出栈顶 / Rising edge: pop top
    bPeek      : BOOL;                     // TRUE：fTop 输出当前栈顶（不改变栈） / TRUE: expose top without popping
    bClear     : BOOL;                     // TRUE：清空栈与锁存（保留累计计数） / TRUE: clear stack and latches, counters kept
    bEnable    : BOOL := TRUE;             // 使能，FALSE 时禁止入栈/出栈 / Enable, FALSE blocks push and pop
END_VAR
VAR_OUTPUT
    fTop       : LREAL;                    // 栈顶值 [EU]，空栈时为 0.0 哨兵 / Top value [EU], 0.0 sentinel when empty
    fPopValue  : LREAL;                    // 本次弹出值 [EU]，未弹出为 0.0 / Popped value [EU], 0.0 when nothing popped
    nCount     : INT;                      // 当前深度 [个]，值域 0..64 / Current depth [count], range 0..64
    bEmpty     : BOOL;                     // 空栈标志 / Empty flag
    bFull      : BOOL;                     // 满栈标志 / Full flag
    bOverflow  : BOOL;                     // 上溢锁存（压栈被拒） / Overflow latched, push rejected
    bUnderflow : BOOL;                     // 下溢锁存（弹栈被拒） / Underflow latched, pop rejected
    uPushCount : UDINT;                    // 累计入栈次数（饱和），仅成功写入时递增 / Total successful pushes, saturating
    uPopCount  : UDINT;                    // 累计出栈次数（饱和），仅成功弹出时递增 / Total successful pops, saturating
    bError     : BOOL;                     // 故障标志（上溢/下溢锁存） / Fault flag, latched
    uErrorId   : UDINT;                    // 故障码，0 = 无故障 / Error code, 0 = no error
    eState     : E_DL_StackState;          // 当前状态（供诊断） / Current state for diagnostics
END_VAR
VAR
    fbTrigPush : R_TRIG;                   // 压栈沿检测实例 / Push edge detector instance
    fbTrigPop  : R_TRIG;                   // 弹栈沿检测实例 / Pop edge detector instance
    afStack    : ARRAY[0..63] OF LREAL;    // 栈体 [EU] / Stack body [EU]
    nTop       : INT;                      // 栈顶指针 = 元素个数，0 = 空 / Top pointer = element count, 0 = empty
    bOvfLatch  : BOOL;                     // 上溢锁存 / Overflow latch
    bUnfLatch  : BOOL;                     // 下溢锁存 / Underflow latch
    eStateInt  : E_DL_StackState;          // 内部状态机当前态 / Internal state machine state
END_VAR
VAR CONSTANT
    DL_LIFO_CAP     : INT   := 64;           // 栈容量，必须与数组维度严格一致 / Capacity, must match the array
    DL_LIFO_CNT_MAX : UDINT := 16#FFFF_FFFE; // 累计计数饱和值，不回绕 / Counter saturation, no wrap-around
END_VAR

(*------------------------------------------------------------------------------
 * 段 1｜无条件刷新区（红线 R7）：两个边沿实例位于主体最前部，严禁进入 IF / CASE
 *      Unconditional refresh zone: both edge instances run at the very top
 *-----------------------------------------------------------------------------*)
fbTrigPush(CLK := bPush);
fbTrigPop(CLK  := bPop);

(*------------------------------------------------------------------------------
 * 段 2｜弹出值本周期清零（边界 B2）：未弹出时输出 0.0 哨兵而非保留上次值，
 *      Popped value cleared every scan
 *      保留上次值会让调用方把旧数据当新数据用
 *-----------------------------------------------------------------------------*)
fPopValue := 0.0;

(*------------------------------------------------------------------------------
 * 段 3｜清空（边界 B5）：电平触发、最高优先级，先于压弹处理；
 *      Clear: level-triggered, highest priority, handled before push and pop
 *      bClear 是唯一清锁存路径；累计计数为生命周期统计，不清零
 *-----------------------------------------------------------------------------*)
IF bClear THEN
    nTop      := 0;
    bOvfLatch := FALSE;
    bUnfLatch := FALSE;
    uErrorId  := 16#0000_0000;
    fTop      := 0.0;
END_IF

(*------------------------------------------------------------------------------
 * 段 4｜压栈（边界 B1/B4）：满栈拒绝写入，绝不覆盖栈底；
 *      Push: rejected when full, the deepest element is never overwritten
 *      拒绝路径不递增累计计数，避免"溢出一次计数暴涨"（边界 B4）
 *-----------------------------------------------------------------------------*)
IF fbTrigPush.Q AND bEnable THEN

    IF nTop >= DL_LIFO_CAP THEN
        bOvfLatch := TRUE;
        uErrorId  := 16#0001_0009;      // 上溢：满栈压入被拒 / Overflow: push rejected on full stack
    ELSIF (nTop >= 0) AND (nTop < DL_LIFO_CAP) THEN
        (* 栈顶指针双检（红线 R4）：写入前显式校验上下界 *)
        (* Top pointer double check: explicit bounds check before writing *)
        afStack[nTop] := fPushValue;
        nTop := nTop + 1;
        IF uPushCount < DL_LIFO_CNT_MAX THEN
            uPushCount := uPushCount + 1;
        END_IF
    ELSE
        (* 指针异常兜底：正常流程不可达，命中说明内存被外部破坏 *)
        (* Pointer anomaly fallback: unreachable in normal flow, memory corruption *)
        bOvfLatch := TRUE;
        uErrorId  := 16#0001_0007;      // 栈顶指针越界 / Top pointer out of range
    END_IF

END_IF

(*------------------------------------------------------------------------------
 * 段 5｜弹栈（边界 B2/B3）：空栈拒绝，弹出值置 0.0 哨兵；
 *      Pop: rejected when empty, popped value set to the 0.0 sentinel
 *      与压栈同周期出现时按"先压后弹"处理，此处已位于压栈之后（边界 B3）
 *-----------------------------------------------------------------------------*)
IF fbTrigPop.Q AND bEnable THEN

    IF nTop <= 0 THEN
        bUnfLatch := TRUE;
        uErrorId  := 16#0001_000A;      // 下溢：空栈弹出被拒 / Underflow: pop rejected on empty stack
        fPopValue := 0.0;
    ELSE
        nTop := nTop - 1;
        IF (nTop >= 0) AND (nTop < DL_LIFO_CAP) THEN
            (* 读回前下标双检（红线 R4） *)
            (* Index double check before read-back *)
            fPopValue := afStack[nTop];
        ELSE
            fPopValue := 0.0;
            uErrorId  := 16#0001_0007;  // 栈顶指针越界 / Top pointer out of range
        END_IF
        IF uPopCount < DL_LIFO_CNT_MAX THEN
            uPopCount := uPopCount + 1;
        END_IF
    END_IF

END_IF

(*------------------------------------------------------------------------------
 * 段 6｜状态派生：锁存优先，其次按深度分空/就绪
 *      State derivation: latches first, then empty or ready by depth
 *-----------------------------------------------------------------------------*)
IF bOvfLatch OR bUnfLatch THEN
    eStateInt := E_DL_StackState.eFault;
ELSIF nTop <= 0 THEN
    eStateInt := E_DL_StackState.eEmpty;
ELSE
    eStateInt := E_DL_StackState.eReady;
END_IF

(*------------------------------------------------------------------------------
 * 段 7｜主状态机（红线 R6）：ENUM + CASE + ELSE 兜底
 *      Main state machine with ELSE fallback
 *      故障态仍允许反向操作（满栈可弹、空栈可压），仅置故障标志（见规格语义表）
 *-----------------------------------------------------------------------------*)
CASE eStateInt OF

    E_DL_StackState.eEmpty:
        (* 空栈：栈顶输出哨兵 0.0 / Empty: top outputs the 0.0 sentinel *)
        fTop := 0.0;

    E_DL_StackState.eReady:
        (* 就绪：栈顶输出 afStack[nTop-1]，读前下标双检（红线 R4） *)
        (* Ready: top outputs afStack[nTop-1] with a bounds check before read *)
        IF (nTop > 0) AND (nTop <= DL_LIFO_CAP) THEN
            fTop := afStack[nTop - 1];
        ELSE
            fTop := 0.0;
        END_IF

    E_DL_StackState.eFault:
        (* 故障锁存：保持现状，bClear 在段 3 解除 / Fault latched, cleared via bClear *)

    ELSE
        (* 非法状态一律回故障态并置码（红线 R6） *)
        (* Illegal state falls back to fault with a code *)
        eStateInt := E_DL_StackState.eFault;
        uErrorId  := 16#0001_0005;

END_CASE

(*------------------------------------------------------------------------------
 * 段 8｜输出单一出口：空满标志由指针派生，指针只在成功路径上增减
 *      Single output exit: flags derived from the pointer, which only moves on success
 *-----------------------------------------------------------------------------*)
nCount     := nTop;
bEmpty     := (nTop <= 0);
bFull      := (nTop >= DL_LIFO_CAP);
bOverflow  := bOvfLatch;
bUnderflow := bUnfLatch;
bError     := (bOvfLatch OR bUnfLatch);
eState     := eStateInt;
END_FUNCTION_BLOCK

(* ---- FB_DL_MedianFilter.st ---- *)
(*==============================================================================
 * 组件名称 (Component)  : FB_DL_MedianFilter
 * 所属子库 (Sublibrary) : DL_MathData
 * 当前版本 (Version)    : 1.0.0
 * 兼容性   (Platform)   : CODESYS 3.5 / TwinCAT 3 / 汇川 InoProShop / Machine Expert
 *                         仅依赖 Standard.library（ABS / MIN / MOD），无厂商方言
 * 功能描述 (Function)   : 滑动窗口中值滤波器（窗口 3..15，强制奇数）。
 *                         对孤立脉冲干扰（变频器干扰、接触器拉弧、单次 AD 跳变）
 *                         免疫：窗口内 1 个坏点被整体剔除，而均值滤波会把坏点
 *                         摊到全窗。用于称重、温度、压力、位置反馈的采集前端。
 *                         启动阶段不等装满：输出"已到样本"的中值，保证上电即有
 *                         合理值，避免 PID 把启动期 0 误认为测量值而满输出。
 * 本文件内含       : E_DL_MedianState（枚举，归属本组件）
 *                    FB_DL_MedianFilter（功能块主体）
 * 开源溯源 (Origin)     : 原创实现（参考西门子 LGF 测量评估组的滤波器分类方式
 *                         与 OSCAT Basic 中值函数"排序后取中"的行为定义
 *                         （EPL-2.0）；OSCAT 采用地址指针入参且会原地排序传入
 *                         数组，本块改为内部副本排序、无指针、无副作用，
 *                         clean-room 编写，未复制任何源码）。
 * 依赖     (Depends)    : 无 DL_ 内部依赖
 * 红线自检 (Redline)    : R1 ✓ 零全局变量表与外部变量引用 ｜ R2 ✓ 零物理 IO 地址直写
 *                         R3 ✓ 纯 IEC 61131-3，无位访问方言与私有指令
 *                         R4 ✓ 窗口钳位 + 环形取数正数化取模 + 下标双检 + NaN 跳过
 *                         R5 ✓ 全变量中英双语同行注释 ｜ R6 ✓ ENUM + CASE + ELSE 兜底
 *                         R7 N/A（无定时器/边沿实例）
 *
 * 【排序副本披露 / Sorting-copy disclosure（边界 B4）】
 *   排序在副本 afSort 上进行，绝不原地排序环形窗 afWindow——
 *   原地排序会打乱环形时间顺序，后续取"最近 N 个样本"时取到错值。
 *
 * 【环形回退取数 / Ring look-back（边界 B3）】
 *   取最近样本用 (写指针 - 1 - k + 容量×2) 取模：先加两倍容量再取模，
 *   把被减数正数化，规避负数取模的跨平台行为差异。
 *
 * 【偶数窗口 / Even window（边界 B2）】
 *   偶数窗口无唯一中值，强制加 1 变奇数，绝不静默取"中间两个的平均"
 *   ——那会退化成均值，尖峰重新渗入输出。
 *
 * 【选型公式 / Sizing formula（边界 B6）】
 *   中值只剔除孤立尖峰。若干扰持续 ≥ 半个窗口宽度，中值仍会被带偏；
 *   窗口长度应 ≥ 2 × 干扰持续采样数 + 1。
 * 【验收向量 / Acceptance vectors】
 *   V1  窗口 5，序列 10,11,10,100,10 → 装满后 fMedian = 10（100 被剔除；
 *       同序列均值 = 28.2，对比可见中值的抗尖峰价值）
 *   V2  窗口 5，仅采 10,10,10 → nFilled = 3、fMedian = 10、eFilling（上电即有值）
 *   V3  窗口 5，采 1,2,3,4,5 → fMedian = 3
 *   V4  窗口设 4（偶数）→ 生效 5、uErrorId = 16#0001_0001
 *   V5  V3 后窗口改为 3 → 整窗重填（nFilled 归 0 再累）、16#0001_0001
 *   V6  bClear 一拍 → nFilled = 0、bValid = FALSE
 * 修订历史 (Revision)   :
 *   2026-11-14  v1.0.0  首版入库（Phase 1 收口批次 · R3）
 *============================================================================*)
TYPE E_DL_MedianState :
(
    eEmpty   := 0,    // 未采到任何样本 / No samples yet
    eFilling := 10,   // 窗口未满，输出已到样本的中值 / Filling, median of available samples
    eReady   := 20,   // 窗口已满 / Window full
    eFault   := 99    // 参数非法当拍（已钳位，下拍恢复）/ Parameter event scan, clamped, recovers next scan
);
END_TYPE

FUNCTION_BLOCK FB_DL_MedianFilter
VAR_INPUT
    fIn       : REAL;                      // 采样输入 [EU] / Sample input [EU]
    bSample   : BOOL := TRUE;              // TRUE = 本拍采一个样本（给单周期脉冲即按需采样） / TRUE: take one sample this scan
    nWindow   : INT   := 5;                // 窗口长度，奇数 3..15，偶数自动加 1，越界钳位 / Window length, odd 3..15, even forced odd
    bClear    : BOOL;                      // TRUE：清空窗口重新填充 / TRUE: clear window and refill
END_VAR
VAR_OUTPUT
    fMedian   : REAL;                      // 中值输出 [EU] / Median output [EU]
    nFilled   : INT;                       // 当前有效样本数 [个]，0..窗口长 / Valid sample count, 0..window length
    bValid    : BOOL;                      // 至少有 1 个样本 / At least one sample available
    bWindowFull : BOOL;                    // 窗口已满 / Window full flag
    uErrorId  : UDINT;                     // 故障码，0 = 无故障（本块码均为瞬时，逐拍重算） / Error code, transient, recomputed every scan
    eState    : E_DL_MedianState;          // 当前状态（供诊断） / Current state for diagnostics
END_VAR
VAR
    afWindow  : ARRAY[0..14] OF REAL;      // 环形样本窗 [EU] / Circular sample window [EU]
    afSort    : ARRAY[0..14] OF REAL;      // 排序副本（不破坏原窗时间顺序） / Sorting copy, ring order untouched
    nWrite    : INT;                       // 写指针，值域 0..14 / Write index, range 0..14
    nFilledInt: INT;                       // 有效样本数（内部） / Internal valid sample count
    nWinEff   : INT;                       // 生效窗口（钳位与奇数化后） / Effective odd window after clamping
    nLastWin  : INT;                       // 上拍生效窗口（变更检测，触发整窗重填） / Previous effective window, change forces refill
    nI        : INT;                       // 插入排序外层索引 / Insertion sort outer index
    nJ        : INT;                       // 插入排序内层索引 / Insertion sort inner index
    nK        : INT;                       // 环形取数索引 / Ring fetch index
    nIdx      : INT;                       // 环形取数换算下标 / Resolved ring index
    fTmp      : REAL;                      // 插入排序交换临时量 [EU] / Insertion sort swap temp [EU]
    nGuard    : INT;                       // 排序防死锁计数器 / Sort guard counter
    bParamEvt : BOOL;                      // 本拍发生参数钳位或窗口变更 / Parameter clamp or window change this scan
    bShiftEnd : BOOL;                      // 本轮内层回退结束标志 / Inner shift finished flag
    bGuardTrip: BOOL;                      // 守卫超限标志（本拍） / Guard tripped flag this scan
    eStateInt : E_DL_MedianState;          // 内部状态机当前态 / Internal state machine state
END_VAR
VAR CONSTANT
    DL_MED_WIN_MIN : INT   := 3;          // 最小窗口 / Minimum window
    DL_MED_WIN_MAX : INT   := 15;         // 最大窗口（= 数组维度） / Maximum window, equals the array dimension
    DL_MED_CAP     : INT   := 15;         // 环形容量，必须与数组维度严格一致 / Ring capacity, must match the array
    DL_MED_EPS     : REAL  := 1.0E-6;     // 浮点判零容差 / Float zero tolerance
    DL_MED_INF_LIM : REAL  := 1.0E30;     // 非有限值判据阈值（超此视为 Inf） / Infinity threshold for non-finite detection
    DL_MED_GUARD   : INT   := 225;        // 排序循环防死锁上限（容量平方） / Sort guard limit, capacity squared
END_VAR

(*------------------------------------------------------------------------------
 * 段 1｜故障码本周期清零：本块故障码全部为瞬时码，逐拍重算
 *      Error code cleared every scan: all codes are transient
 *-----------------------------------------------------------------------------*)
uErrorId  := 16#0000_0000;
bParamEvt := FALSE;
bGuardTrip:= FALSE;
nGuard    := 0;

(*------------------------------------------------------------------------------
 * 段 2｜窗口规整（边界 B2）：越界钳位、偶数强制奇数，只在本拍置码不刷屏
 *      Window normalization: clamp and force odd, code set only on the event scan
 *-----------------------------------------------------------------------------*)
nWinEff := nWindow;
IF nWinEff < DL_MED_WIN_MIN THEN
    nWinEff  := DL_MED_WIN_MIN;
    bParamEvt := TRUE;
END_IF
IF nWinEff > DL_MED_WIN_MAX THEN
    nWinEff  := DL_MED_WIN_MAX;
    bParamEvt := TRUE;
END_IF
IF (nWinEff MOD 2) = 0 THEN
    nWinEff  := MIN(nWinEff + 1, DL_MED_WIN_MAX);
    bParamEvt := TRUE;
END_IF
IF bParamEvt THEN
    uErrorId := 16#0001_0001;           // 窗口非法已钳位 / Window invalid, clamped
END_IF

(*------------------------------------------------------------------------------
 * 段 3｜窗口变更检测（R14 语义参数变更）：生效窗口与上拍不同 → 整窗作废。
 *      Window change detection: effective window differs, whole window voided
 *      新旧窗口混填的中值无物理意义；重填会有一个窗口长度的空档
 *-----------------------------------------------------------------------------*)
IF nWinEff <> nLastWin THEN
    nFilledInt := 0;
    nWrite     := 0;
    IF nLastWin <> 0 THEN               // 上电首扫不算参数事件 / Power-up first scan is not a parameter event
        uErrorId  := 16#0001_0001;      // 窗口变更触发重填 / Window change forces refill
        bParamEvt := TRUE;
    END_IF
END_IF
nLastWin := nWinEff;

(*------------------------------------------------------------------------------
 * 段 4｜清空：电平触发，先于采样处理
 *      Clear: level-triggered, handled before sampling
 *-----------------------------------------------------------------------------*)
IF bClear THEN
    nFilledInt := 0;
    nWrite     := 0;
END_IF

(*------------------------------------------------------------------------------
 * 段 5｜采样（边界：NaN/Inf 跳过不入窗）
 *      Sampling: NaN or Inf samples are skipped, never stored
 *-----------------------------------------------------------------------------*)
IF bSample THEN
    IF (fIn <> fIn) OR (ABS(fIn) > DL_MED_INF_LIM) THEN
        uErrorId := 16#0001_0006;       // 样本非有限值已跳过 / Non-finite sample skipped
    ELSIF (nWrite >= 0) AND (nWrite < DL_MED_CAP) THEN
        (* 写指针双检（红线 R4）：MOD 已保证范围，仍显式兜底防越界写 *)
        (* Write index double check: explicit guard besides MOD *)
        afWindow[nWrite] := fIn;
        nWrite    := (nWrite + 1) MOD DL_MED_CAP;
        nFilledInt := MIN(nFilledInt + 1, nWinEff);
    END_IF
END_IF

(*------------------------------------------------------------------------------
 * 段 6｜取有效样本到排序副本（边界 B3）：只取最近 nFilledInt 个，
 *      Copy the valid samples into the sorting copy
 *      禁止复制整窗——未填区是 0，会把中值拉低
 *-----------------------------------------------------------------------------*)
FOR nK := 0 TO (nFilledInt - 1) DO
    (* 正数化取模：先加两倍容量再取模，规避负数取模的平台差异（边界 B3） *)
    (* Positive modulo: add twice the capacity before MOD, platform-safe *)
    nIdx := (nWrite - 1 - nK + DL_MED_CAP * 2) MOD DL_MED_CAP;
    IF (nIdx >= 0) AND (nIdx < DL_MED_CAP) AND (nK >= 0) AND (nK < DL_MED_CAP) THEN
        afSort[nK] := afWindow[nIdx];
    END_IF
END_FOR;

(*------------------------------------------------------------------------------
 * 段 7｜插入排序（边界 B4）：对副本 afSort[0..nFilledInt-1] 排序，
 *      Insertion sort on the copy afSort[0..nFilledInt-1]
 *      n ≤ 15 最坏 105 次比较；nGuard 防死锁，超限置 16#0001_0004
 *-----------------------------------------------------------------------------*)
FOR nI := 1 TO (nFilledInt - 1) DO
    fTmp      := afSort[nI];
    nJ        := nI - 1;
    bShiftEnd := FALSE;
    WHILE (nJ >= 0) AND (NOT bShiftEnd) DO
        nGuard := nGuard + 1;
        IF nGuard > DL_MED_GUARD THEN
            uErrorId   := 16#0001_0004; // 排序循环保护触发 / Sort loop guard tripped
            bGuardTrip := TRUE;         // 本拍放弃落位，保留已排部分 / Drop this pass, keep the sorted part
            bShiftEnd  := TRUE;
        ELSIF afSort[nJ] > fTmp THEN
            afSort[nJ + 1] := afSort[nJ];
            nJ := nJ - 1;
        ELSE
            bShiftEnd := TRUE;
        END_IF
    END_WHILE
    IF NOT bGuardTrip THEN
        afSort[nJ + 1] := fTmp;         // 正常路径含 nJ = -1 时落位到队首 / Normal path, nJ = -1 lands at the front
    END_IF
END_FOR;

(*------------------------------------------------------------------------------
 * 段 8｜取中值：奇数取正中；偶数为防御分支（正常流程已被 B2 排除）
 *      Median extraction: odd takes the middle; even is defensive only
 *-----------------------------------------------------------------------------*)
IF nFilledInt > 0 THEN
    IF (nFilledInt MOD 2) = 1 THEN
        fMedian := afSort[nFilledInt / 2];              // 整除取正中 / Integer division takes the middle
    ELSE
        fMedian := (afSort[nFilledInt / 2 - 1] + afSort[nFilledInt / 2]) / 2.0;
    END_IF
ELSE
    fMedian := 0.0;                     // 空窗输出 0.0 哨兵 / Empty window outputs the 0.0 sentinel
END_IF

(*------------------------------------------------------------------------------
 * 段 9｜状态派生与主状态机（红线 R6）：ENUM + CASE + ELSE 兜底
 *      State derivation and main state machine with ELSE fallback
 *-----------------------------------------------------------------------------*)
IF bParamEvt THEN
    eStateInt := E_DL_MedianState.eFault;
ELSIF nFilledInt <= 0 THEN
    eStateInt := E_DL_MedianState.eEmpty;
ELSIF nFilledInt < nWinEff THEN
    eStateInt := E_DL_MedianState.eFilling;
ELSE
    eStateInt := E_DL_MedianState.eReady;
END_IF

CASE eStateInt OF

    E_DL_MedianState.eEmpty:
        (* 空窗：无有效输出，bValid 由段 10 置 FALSE / Empty: no valid output *)

    E_DL_MedianState.eFilling:
        (* 填充中：段 8 已按已到样本取中值，保证上电即有值（边界 B1） *)
        (* Filling: median of available samples, a value from power-up on *)

    E_DL_MedianState.eReady:
        (* 就绪：整窗中值 / Ready: full-window median *)

    E_DL_MedianState.eFault:
        (* 参数事件当拍：参数已修正、下拍恢复，不锁存 / Event scan, recovers next scan *)

    ELSE
        (* 非法状态一律回故障态并置码（红线 R6） *)
        (* Illegal state falls back to fault with a code *)
        eStateInt := E_DL_MedianState.eFault;
        uErrorId  := 16#0001_0005;

END_CASE

(*------------------------------------------------------------------------------
 * 段 10｜输出单一出口：有效性与满窗标志由计数派生
 *      Single output exit: validity and full flags derived from the count
 *-----------------------------------------------------------------------------*)
nFilled     := nFilledInt;
bValid      := (nFilledInt > 0);
bWindowFull := (nFilledInt >= nWinEff);
eState      := eStateInt;
END_FUNCTION_BLOCK
